(* IEC 61131-3 sources: daoli-st-library/DL_Process (part 18) *)

(* ---- FC_DL_TemperEmpiricalHardnessCalc.st ---- *)
(*
  Component : FC_DL_TemperEmpiricalHardnessCalc
  Category  : DL_Process
  Type      : FC
  Complexity: C2
  VERSION   : v1.0.0
  功能      : 回火温度-硬度经验曲线核算：按四点节点表分段线性插值得到基准 HRC，再按含碳量修正，超界双向钳位。
  开源溯源  : 道莅原创 clean-room 自研（无外部代码引用）｜License: MIT
  边界条件  : ① 节点表必须严格升序且首末温差 > 1e-9，否则返回哨兵 -1；
              ② 回火温度超出节点区间时取端点值并置 xClamped，禁外推；
              ③ 含碳量修正量双侧钳位 ±8 HRC，防小样本经验式发散。
*)
FUNCTION FC_DL_TemperEmpiricalHardnessCalc : REAL
VAR_INPUT
    fTemperC    : REAL;               (* 回火温度 [°C] Tempering temperature *)
    afTempKnot  : ARRAY[0..3] OF REAL;(* 节点温度表（升序） [°C] Knot temperatures ascending *)
    afHrcKnot   : ARRAY[0..3] OF REAL;(* 节点硬度表 [HRC] Knot hardness values *)
    fCarbonPct  : REAL;               (* 钢材含碳量 [%] Carbon content *)
END_VAR
VAR_OUTPUT
    fHrc      : REAL;   (* 插值得到的回火硬度 [HRC] Interpolated hardness *)
    fHrcCorr  : REAL;   (* 含碳量修正后的硬度 [HRC] Carbon-corrected hardness *)
    xClamped  : BOOL;   (* 超界钳位标志 [-] Out-of-range clamp flag *)
    xValid    : BOOL;   (* 计算有效性标志 [-] Calculation valid flag *)
END_VAR
VAR CONSTANT
    DL_EPS       : REAL := 1.0E-9;   (* 除零判定容差 [无量纲] Divide-by-zero tolerance *)
    DL_CORR_K    : REAL := 30.0;     (* 含碳量修正斜率 [HRC/%C] Carbon correction slope *)
    DL_CORR_BASE : REAL := 0.40;     (* 含碳量修正基准 [%C] Carbon correction base *)
    DL_CORR_LIM  : REAL := 8.0;      (* 含碳量修正钳位 [HRC] Carbon correction clamp *)
END_VAR
VAR
    nIdx  : INT;    (* 插值段循环下标 [-] Interpolation segment index *)
    nBad  : INT;    (* 节点表非有限计数，0 = 全部有限 [-] Non-finite knot counter *)
    fDen  : REAL;   (* 当前段温度跨度 [°C] Segment temperature span *)
    fCorr : REAL;   (* 含碳量修正量 [HRC] Carbon correction amount *)
END_VAR
(* 出口预置：四出口统一预置 *)
fHrc := 0.0; fHrcCorr := 0.0; xClamped := FALSE; xValid := FALSE; nBad := 0;
(* 非有限拦截：标量输入自反判 NaN，自身差值判 Inf *)
IF (fTemperC <> fTemperC) OR ((fTemperC - fTemperC) <> 0.0)
   OR (fCarbonPct <> fCarbonPct) OR ((fCarbonPct - fCarbonPct) <> 0.0) THEN
    FC_DL_TemperEmpiricalHardnessCalc := -1.0;  (* 哨兵 -1：输入非有限 / Sentinel -1 non-finite *)
    RETURN;
END_IF
(* 节点表非有限拦截：四个温度节点与四个硬度节点逐个判（越界读前先判界） *)
FOR nIdx := 0 TO 3 DO
    IF (nIdx >= 0) AND (nIdx <= 3) THEN
        IF (afTempKnot[nIdx] <> afTempKnot[nIdx])
           OR ((afTempKnot[nIdx] - afTempKnot[nIdx]) <> 0.0)
           OR (afHrcKnot[nIdx] <> afHrcKnot[nIdx])
           OR ((afHrcKnot[nIdx] - afHrcKnot[nIdx]) <> 0.0) THEN
            nBad := nBad + 1;
        END_IF
    END_IF
END_FOR
IF nBad > 0 THEN
    FC_DL_TemperEmpiricalHardnessCalc := -1.0;  (* 哨兵 -1：节点表非有限 / Sentinel -1 bad knots *)
    RETURN;
END_IF
(* 节点表域闸：首末温差必须为正，保证区间可插值与升序约定 *)
IF (afTempKnot[3] - afTempKnot[0]) <= DL_EPS THEN
    FC_DL_TemperEmpiricalHardnessCalc := -1.0;  (* 哨兵 -1：节点表非法 / Sentinel -1 bad knot table *)
    RETURN;
END_IF
(* 超界钳位：低于首节点取首值，高于末节点取末值，禁外推 *)
IF fTemperC <= afTempKnot[0] THEN
    fHrc := afHrcKnot[0];                       (* 端点取值 [HRC] / Lower endpoint *)
    xClamped := TRUE;                           (* 低位钳位标志 [-] / Low clamp *)
ELSIF fTemperC >= afTempKnot[3] THEN
    fHrc := afHrcKnot[3];                       (* 端点取值 [HRC] / Upper endpoint *)
    xClamped := TRUE;                           (* 高位钳位标志 [-] / High clamp *)
ELSE
    (* 分段线性插值：升序镜像遍历（禁倒序循环关键字），下标上限 2 保证 i+1 <= 3 不越界 *)
    FOR nIdx := 0 TO 2 DO
        IF (fTemperC >= afTempKnot[nIdx]) AND (fTemperC <= afTempKnot[nIdx + 1]) THEN
            fDen := afTempKnot[nIdx + 1] - afTempKnot[nIdx];   (* 段跨度 [°C] / Segment span *)
            IF ABS(fDen) > DL_EPS THEN
                fHrc := afHrcKnot[nIdx]
                        + (afHrcKnot[nIdx + 1] - afHrcKnot[nIdx])
                          * (fTemperC - afTempKnot[nIdx]) / fDen;
            END_IF
        END_IF
    END_FOR
END_IF
(* 含碳量修正：以 0.40 %C 为基准，每 0.1 %C 约 3 HRC，双侧钳位 *)
fCorr := (fCarbonPct - DL_CORR_BASE) * DL_CORR_K;
IF fCorr > DL_CORR_LIM THEN
    fCorr := DL_CORR_LIM;                       (* 上限钳位 [HRC] / Upper clamp *)
ELSIF fCorr < -DL_CORR_LIM THEN
    fCorr := -DL_CORR_LIM;                      (* 下限钳位 [HRC] / Lower clamp *)
END_IF
fHrcCorr := fHrc + fCorr;                       (* 修正后硬度 [HRC] / Corrected hardness *)
xValid := TRUE;                                 (* 链路有效 / Chain valid *)
FC_DL_TemperEmpiricalHardnessCalc := fHrcCorr;  (* 返回修正硬度 [HRC] / Return hardness *)
END_FUNCTION

(* ---- FC_DL_ThickenerSettlingAreaCalc.st ---- *)
(*
  Name: FC_DL_ThickenerSettlingAreaCalc
  Category: DL_Process
  Version: 1.0.0
  Round: R89 / 2026-11-25
  开源溯源：clean-room 自研（族 矿山破碎筛分，ST 开源生态实测 0 命中，无外部代码引入）
  功能：按固体体积衡算求浓密机底流体积流量与溢流量，再用沉降速度法算所需沉降面积与上升流速。
  边界条件：① 四入参全部过非有限闸，任一非有限返回哨兵 -1；
            ② 底流浓度必须显著高于给矿浓度（差值 ≥ 1 %），否则衡算无解，返回哨兵 -1；
            ③ 体积分数 φ 由质量分数与固/液密度反算，分母（固相项 + 液相项）在 0~1 质量分数域内恒正，
               仍以 DL_EPS 兜底防浮点下溢；面积取安全系数 1.15，上升流速 = Qo/A 故恒低于沉降速度。
  量纲自证：Q[m3/h] ÷ v[m/h] = m2；φ 无量纲。
*)
FUNCTION FC_DL_ThickenerSettlingAreaCalc : REAL
VAR_INPUT
    fFeedM3h : REAL;         (* 给矿浆体流量 [m3/h] Feed slurry flow [m3/h] *)
    fFeedSolidsPct : REAL;   (* 给矿固体质量浓度 [%] Feed solids mass concentration [%] *)
    fUnderSolidsPct : REAL;  (* 底流固体质量浓度 [%] Underflow solids mass concentration [%] *)
    fSettlingVel : REAL;     (* 自由沉降速度 [m/h] Free settling velocity [m/h] *)
END_VAR
VAR_OUTPUT
    fAreaM2 : REAL;          (* 所需沉降面积（含安全系数） [m2] Required settling area [m2] *)
    fRiseVel : REAL;         (* 溢流上升流速 [m/h] Overflow rise velocity [m/h] *)
    fOverflowM3h : REAL;     (* 溢流浆体流量 [m3/h] Overflow flow [m3/h] *)
    xSizingOk : BOOL;        (* 上升流速低于沉降速度则 TRUE [-] Rise velocity below settling velocity *)
    xValid : BOOL;           (* 计算有效性标志 [-] Calculation valid flag *)
END_VAR
VAR CONSTANT
    DL_EPS : REAL := 1.0E-9;      (* 除零判定容差 [-] Divide-by-zero tolerance *)
    DL_RHO_S : REAL := 2.7;       (* 固体密度（矿浆通用取值） [t/m3] Solids density [t/m3] *)
    DL_RHO_W : REAL := 1.0;       (* 液相密度（水） [t/m3] Liquid density [t/m3] *)
    DL_SF : REAL := 1.15;         (* 面积安全系数 [-] Area safety factor *)
    DL_PCT : REAL := 100.0;       (* 百分数基准 [%] Percent base *)
    DL_CONC_MIN_DIFF : REAL := 1.0; (* 底流与给矿浓度最小差值 [%] Minimum concentration difference *)
END_VAR
VAR
    fCf : REAL;     (* 给矿质量分数 [-] Feed mass fraction *)
    fCu : REAL;     (* 底流质量分数 [-] Underflow mass fraction *)
    fPhiF : REAL;   (* 给矿固体体积分数 [-] Feed solids volume fraction *)
    fPhiU : REAL;   (* 底流固体体积分数 [-] Underflow solids volume fraction *)
    fQs : REAL;     (* 固体体积流量 [m3/h] Solids volume flow [m3/h] *)
    fQu : REAL;     (* 底流浆体体积流量 [m3/h] Underflow slurry flow [m3/h] *)
    fQo : REAL;     (* 溢流浆体体积流量 [m3/h] Overflow flow [m3/h] *)
END_VAR
(* 出口预置：五出口统一预置（R256） *)
fAreaM2 := 0.0; fRiseVel := 0.0; fOverflowM3h := 0.0; xSizingOk := FALSE; xValid := FALSE;
(* 非有限闸：NaN 自反判 + Inf 差值自减判，四入参全枚举（R272） *)
IF (fFeedM3h <> fFeedM3h) OR ((fFeedM3h - fFeedM3h) <> 0.0)
   OR (fFeedSolidsPct <> fFeedSolidsPct) OR ((fFeedSolidsPct - fFeedSolidsPct) <> 0.0)
   OR (fUnderSolidsPct <> fUnderSolidsPct) OR ((fUnderSolidsPct - fUnderSolidsPct) <> 0.0)
   OR (fSettlingVel <> fSettlingVel) OR ((fSettlingVel - fSettlingVel) <> 0.0) THEN
    FC_DL_ThickenerSettlingAreaCalc := -1.0;    (* 哨兵 -1：入参非有限 / Sentinel -1, non-finite input *)
    RETURN;
END_IF
(* 组态域闸：流量与沉降速度为除子，浓度须物理可行且底流显著高于给矿 *)
IF (fFeedM3h <= DL_EPS) OR (fSettlingVel <= DL_EPS)
   OR (fFeedSolidsPct <= 0.0) OR (fFeedSolidsPct >= DL_PCT)
   OR (fUnderSolidsPct <= 0.0) OR (fUnderSolidsPct > DL_PCT)
   OR ((fUnderSolidsPct - fFeedSolidsPct) < DL_CONC_MIN_DIFF) THEN
    FC_DL_ThickenerSettlingAreaCalc := -1.0;    (* 哨兵 -1：组态非法 / Sentinel -1, bad configuration *)
    RETURN;
END_IF
fCf := fFeedSolidsPct / DL_PCT;                 (* 质量分数 [-] Mass fraction *)
fCu := fUnderSolidsPct / DL_PCT;
(* 体积分数：φ = (C/ρs) / (C/ρs + (1−C)/ρw)，固液体积可加性假设 *)
IF ((fCf / DL_RHO_S) + ((1.0 - fCf) / DL_RHO_W)) <= DL_EPS THEN
    FC_DL_ThickenerSettlingAreaCalc := -1.0;    (* 哨兵 -1：体积分数塌零 / Sentinel -1, vanishing phi *)
    RETURN;
END_IF
fPhiF := (fCf / DL_RHO_S) / ((fCf / DL_RHO_S) + ((1.0 - fCf) / DL_RHO_W));
fPhiU := (fCu / DL_RHO_S) / ((fCu / DL_RHO_S) + ((1.0 - fCu) / DL_RHO_W));
(* 固体体积衡算：Qs = Qf·φf；底流体积 Qu = Qs/φu，φu 已过域闸恒正 *)
IF fPhiU <= DL_EPS THEN
    FC_DL_ThickenerSettlingAreaCalc := -1.0;    (* 哨兵 -1：底流体积分数塌零 / Sentinel -1, phi underflow zero *)
    RETURN;
END_IF
fQs := fFeedM3h * fPhiF;                        (* 固体体积流量 [m3/h] Solids volume flow *)
fQu := fQs / fPhiU;                             (* 底流浆体流量 [m3/h] Underflow slurry flow *)
fQo := fFeedM3h - fQu;                          (* 溢流 = 给矿 − 底流 [m3/h] Overflow flow *)
IF fQo <= DL_EPS THEN
    FC_DL_ThickenerSettlingAreaCalc := -1.0;    (* 哨兵 -1：衡算无溢流，组态矛盾 / Sentinel -1, no overflow *)
    RETURN;
END_IF
(* 沉降面积：A = Qo/v × SF，Qo[m3/h] ÷ v[m/h] = m2 *)
fAreaM2 := (fQo / fSettlingVel) * DL_SF;
(* 上升流速：vR = Qo/A，A 已过正性检查（上式保证 ≥ SF 倍正量） *)
IF fAreaM2 <= DL_EPS THEN
    FC_DL_ThickenerSettlingAreaCalc := -1.0;    (* 哨兵 -1：面积塌零 / Sentinel -1, vanishing area *)
    RETURN;
END_IF
fRiseVel := fQo / fAreaM2;
fOverflowM3h := fQo;
(* 校核：上升流速低于自由沉降速度（含安全系数后恒成立，此处照实判定） *)
xSizingOk := fRiseVel < fSettlingVel;
xValid := TRUE;                                 (* 链路有效 / Chain valid *)
FC_DL_ThickenerSettlingAreaCalc := fAreaM2;
END_FUNCTION

(* ---- FC_DL_TinBathAtmosphereCalc.st ---- *)
(*
  Name: FC_DL_TinBathAtmosphereCalc
  Category: DL_Process
  Version: 1.0.0
  Round: R90 / 2026-11-25
  开源溯源：clean-room 自研（族 浮法玻璃锡槽退火，ST 开源生态实测 0 命中，无外部代码引入）
  功能：1) 锡槽保护气 H2 配比按「氢耗氧化学计量」估算。漏入锡槽的空气带入氧气，
           氧气与氢按 2H2 + O2 → 2H2O 反应，故 1 体积氧气需要 2 体积氢气中和。
           逐步为：
             氧带入量 = 漏入空气量 × 空气中氧体积分数(0.21)
             需中和氧量 = 氧带入量 − 允许残氧量（目标 ppm 折算为体积流量）
             氢需求 = 2 × 需中和氧量 × 过量系数
             氢配比 = 氢需求 / 保护气总流量 × 100
           允许残氧量按「目标 ppm × 总流量 × 1e-6」折算，使得目标越严格所需氢越多，方向正确。
        2) 过量系数 DL_HSF(1.5) 用于覆盖反应不完全与局部湍流死区，是安全冗余而非效率系数。
  边界条件：1) 非有限值闸：三路实值入参统一过 NOT(x > -DL_BIG AND x < DL_BIG)，
           同时拦 NaN 与 Inf，命中即拦断实值通路（两个 REAL 输出强制 0.0）并置无效（R19）。
        2) 分母零闸：ABS(fTotalFlowM3h) > DL_EPS 才允许算配比（总流量为 0 时配比无定义）。
        3) 负值闸：漏入量、目标氧含量、总流量任一为负判无效（不取绝对值掩盖反向）。
        4) 配比饱和钳制：H2 配比钳 0 ~ DL_H2_MAX(10 %)。上限的依据是保护气进入爆炸下限区间
           （H2 在空气中的爆炸下限约 4 %，但锡槽内为氮基气氛且需维持正压，工艺上按 10 % 上限组态），
           超过上限必须由安全联锁处理，本件只做钳制与无效标记，不做安全切断。
        5) 需求为负（残氧目标高于带入氧）时氢需求钳 0，属合法工况（无需加氢），不判无效。
        6) 饱和钳制：氢流量钳 0 ~ DL_H2_FLOW_MAX(10000 m3/h)，防溢出。
  量纲自证：氧带入量 = (m3/h) × [-] = m3/h；残氧量 = ppm × (m3/h) × 1E-6 = m3/h；
           需中和氧量 = (m3/h) − (m3/h) = m3/h，减法同量纲；
           氢需求 = [-] × (m3/h) × [-] = m3/h（化学计量比与过量系数均为无因次）；
           配比 = (m3/h) / (m3/h) × 100 = 无因次 [%]，分母与分子同量纲。
*)

FUNCTION FC_DL_TinBathAtmosphereCalc : BOOL
VAR_INPUT
    fO2TargetPpm   : REAL;   // 目标残氧含量 [ppm] / Target residual oxygen [ppm]
    fLeakM3h       : REAL;   // 漏入锡槽的空气量 [m3/h] / Air leakage into tin bath [m3/h]
    fTotalFlowM3h  : REAL;   // 保护气总流量 [m3/h] / Total protective gas flow [m3/h]
END_VAR
VAR_OUTPUT
    fH2Pct         : REAL;   // 氢气体积配比 [%] / Hydrogen volume ratio [%]
    fFlowM3h       : REAL;   // 氢气需求体积流量 [m3/h] / Hydrogen required volumetric flow [m3/h]
    xValid         : BOOL;   // 计算有效标志 [bool] / Calculation valid flag [bool]
END_VAR
VAR
    _fO2IngressM3h : REAL;   // 漏入氧气量 [m3/h] / Oxygen ingress [m3/h]
    _fO2AllowM3h   : REAL;   // 允许残氧量 [m3/h] / Allowable residual oxygen [m3/h]
    _fO2NeedM3h    : REAL;   // 需中和氧量 [m3/h] / Oxygen to be neutralized [m3/h]
    _fH2NeedM3h    : REAL;   // 氢需求（含过量系数）[m3/h] / Hydrogen demand with safety factor [m3/h]
    _fPctRaw       : REAL;   // 未饱和的配比 [%] / Raw ratio [%]
END_VAR
VAR CONSTANT
    DL_EPS         : REAL := 1.0E-9;    // 分母零闸阈值 [-] / Division-zero gate threshold [-]
    DL_BIG         : REAL := 1.0E12;    // 非有限值闸量级上限 [-] / Finiteness gate magnitude [-]
    DL_PCT         : REAL := 100.0;     // 百分比换算因子 [%] / Percent conversion factor [%]
    DL_O2_AIR_FRAC : REAL := 0.21;      // 空气中氧体积分数 [-] / Oxygen volume fraction in air [-]
    DL_H2_STOICH   : REAL := 2.0;       // 2H2 + O2 化学计量比 [-] / Hydrogen to oxygen stoichiometry [-]
    DL_PPM_FRAC    : REAL := 1.0E-6;    // ppm → 体积分数换算因子 [-] / ppm to volume fraction factor [-]
    DL_HSF         : REAL := 1.5;       // 氢过量系数（安全冗余）[-] / Hydrogen excess factor [-]
    DL_H2_MAX      : REAL := 10.0;      // 氢配比饱和上限 [%] / Hydrogen ratio saturation ceiling [%]
    DL_H2_FLOW_MAX : REAL := 10000.0;   // 氢流量饱和上限 [m3/h] / Hydrogen flow saturation ceiling [m3/h]
END_VAR

(* —— 段 1：非有限值闸（R19：三路入参全覆盖，拦 NaN 与 Inf） —— *)
IF NOT (fO2TargetPpm > -DL_BIG AND fO2TargetPpm < DL_BIG)
   OR NOT (fLeakM3h > -DL_BIG AND fLeakM3h < DL_BIG)
   OR NOT (fTotalFlowM3h > -DL_BIG AND fTotalFlowM3h < DL_BIG) THEN
    fH2Pct := 0.0;                          // 输出强制 0.0 / Output forced to zero
    fFlowM3h := 0.0;                        // 氢流量强制 0.0 / Hydrogen flow forced to zero
    xValid := FALSE;                        // 有效位清零 / Validity cleared
    FC_DL_TinBathAtmosphereCalc := FALSE;   // 返回码同源 / Return mirrors validity
    RETURN;                                 // 立即退出 / Immediate exit
END_IF

(* —— 段 2：分母零闸（R4：总流量是配比分母） —— *)
IF ABS(fTotalFlowM3h) <= DL_EPS THEN
    fH2Pct := 0.0;                          // 输出强制 0.0 / Output forced to zero
    fFlowM3h := 0.0;                        // 氢流量强制 0.0 / Hydrogen flow forced to zero
    xValid := FALSE;                        // 判无效 / Invalid
    FC_DL_TinBathAtmosphereCalc := FALSE;   // 返回码同步 / Return synchronised
    RETURN;                                 // 提前退出 / Early exit
END_IF

(* —— 段 3：负值闸（漏入量、目标氧含量、总流量均不可为负） —— *)
IF (fO2TargetPpm < 0.0) OR (fLeakM3h < 0.0) OR (fTotalFlowM3h < 0.0) THEN
    fH2Pct := 0.0;                          // 输出强制 0.0 / Output forced to zero
    fFlowM3h := 0.0;                        // 氢流量强制 0.0 / Hydrogen flow forced to zero
    xValid := FALSE;                        // 判无效 / Invalid
    FC_DL_TinBathAtmosphereCalc := FALSE;   // 返回码同步 / Return synchronised
    RETURN;                                 // 提前退出 / Early exit
END_IF

(* —— 段 4：氧衡算（R22 方向自核：漏入氧减去允许残氧，才是需要中和的量） —— *)
_fO2IngressM3h := fLeakM3h * DL_O2_AIR_FRAC;                      // 漏入氧气 [m3/h]
_fO2AllowM3h := fO2TargetPpm * DL_PPM_FRAC * fTotalFlowM3h;       // 允许残氧 [m3/h]
_fO2NeedM3h := MAX(0.0, _fO2IngressM3h - _fO2AllowM3h);           // 需中和氧量 [m3/h]（负值钳 0）

(* —— 段 5：氢需求与配比（化学计量比 2、过量系数 1.5 均为无因次） —— *)
_fH2NeedM3h := DL_H2_STOICH * _fO2NeedM3h * DL_HSF;               // 氢需求 [m3/h]
_fPctRaw := _fH2NeedM3h / fTotalFlowM3h * DL_PCT;                 // 氢配比 [%]

(* —— 段 6：输出单点写盘（饱和钳制） —— *)
fFlowM3h := LIMIT(0.0, _fH2NeedM3h, DL_H2_FLOW_MAX);              // 氢流量 [m3/h]
fH2Pct := LIMIT(0.0, _fPctRaw, DL_H2_MAX);                        // 氢配比 [%]

(* —— 段 7：有效位单点聚合（分母为正 + 入参非负） —— *)
xValid := (fTotalFlowM3h > DL_EPS)                                // 总流量为正
          AND (fO2TargetPpm >= 0.0)                               // 目标残氧非负
          AND (fLeakM3h >= 0.0);                                  // 漏入量非负
FC_DL_TinBathAtmosphereCalc := xValid;                            // 返回码：TRUE = 计算可信

END_FUNCTION

(* ---- FC_DL_TireCureBladderSteamCalc.st ---- *)
(*
  Name: FC_DL_TireCureBladderSteamCalc
  Category: DL_Process
  Version: 1.0.0
  Round: R91 / 2026-11-25
  开源溯源：clean-room 自研（族 轮胎硫化，ST 开源生态实测 0 命中，无外部代码引入）
  功能：1) 单周期胶囊蒸汽耗量按「充装量 + 升温量 + 排凝损失」三段求和：
           充装量 = 胶囊容积 * 蒸汽密度；
           升温量 = 胶囊内容物质量 * 比热 * 温升 / 潜热（把显热需求折成蒸汽质量）；
           排凝损失 = (充装量 + 升温量) * fDrainPct / 100。
           即 m = (V*rho + m*cp*dT/hfg) * (1 + drainPct/100)，单位 kg/周期。
        2) 输出分解量 fFillKg 与 fHeatUpKg，便于按段归因能耗（充装段与升温段的节能措施完全不同）。
        3) 容积零闸与潜热零闸：胶囊容积为充装量的乘子、潜热为升温量的分母，
           任一为零会把「未组态」伪装成「零耗量」，必须判无效而非输出 0。
  边界条件：1) 非有限值闸：七路实值入参先过 NOT(x > -DL_BIG AND x < DL_BIG)，同时拦 NaN 与 Inf，
           命中即闸断实值通路（三段耗量与总耗量强制 0.0），不得只置标志（R19）。
        2) 分母零闸：升华/汽化潜热 fLatentKjKg 必须 > DL_EPS；胶囊内容物比热 fWaterCpKjKgK 必须 > DL_EPS。
        3) 容积零闸：fBladderVolL 必须 > DL_EPS；蒸汽密度 fSteamDensityKgm3 必须 > DL_EPS。
        4) 排凝率域闸：fDrainPct 必须落在 [0.0, DL_DRAIN_HI] 内（排凝率超 100 % 不具物理意义），
           越域判无效不钳制。
        5) 判据取原始值（R24）：总量越域判定使用钳制前的 _fTotalRawKg，钳制只作用于输出。
        6) 纯函数无状态：单周期耗量的累计与班产统计由上层计量模块承担。
  量纲自证：V [L] * rho [kg/m3] / 1000 [L/m3] = kg；
           m [kg] * cp [kJ/(kg*K)] * dT [K] = kJ；kJ / hfg [kJ/kg] = kg；
           三段同为 kg，求和合法；排凝率为无因次百分数，乘 kg 仍为 kg。
  修订历史 Revision :
    2026-11-25  v1.0.0  R91 首版
*)

FUNCTION FC_DL_TireCureBladderSteamCalc : BOOL
VAR_INPUT
    fBladderVolL     : REAL;   // 胶囊有效容积 [L] / Effective bladder volume [L]
    fSteamDensityKgm3 : REAL;  // 工作压力下蒸汽密度 [kg/m3] / Steam density at working pressure [kg/m3]
    fContentMassKg   : REAL;   // 胶囊内容物（水/氮）质量 [kg] / Bladder content mass [kg]
    fWaterCpKjKgK    : REAL;   // 内容物比热 [kJ/(kg*K)] / Content specific heat [kJ/(kg*K)]
    fTempRiseK       : REAL;   // 升温幅度 [K] / Temperature rise [K]
    fLatentKjKg      : REAL;   // 工作压力下汽化潜热 [kJ/kg] / Latent heat of vaporisation [kJ/kg]
    fDrainPct        : REAL;   // 排凝损失占充装与升温之和的百分比 [%] / Blowdown loss percentage [%]
END_VAR
VAR_OUTPUT
    fFillKg          : REAL;   // 充装段蒸汽量 [kg] / Steam for initial filling [kg]
    fHeatUpKg        : REAL;   // 升温段蒸汽量 [kg] / Steam for heat-up [kg]
    fSteamKg         : REAL;   // 单周期蒸汽总耗量 [kg/cycle] / Total steam consumption per cycle [kg/cycle]
    xValid           : BOOL;   // 计算有效标志 [bool] / Calculation valid flag [bool]
END_VAR
VAR
    _fFillRawKg      : REAL;   // 钳制前的充装量 [kg] / Raw fill mass [kg]
    _fHeatRawKg      : REAL;   // 钳制前的升温量 [kg] / Raw heat-up mass [kg]
    _fTotalRawKg     : REAL;   // 钳制前的总量 [kg] / Raw total mass [kg]
    _fDrainFactor    : REAL;   // 排凝放大因子（1 + 排凝率/100）[-] / Blowdown multiplier [-]
END_VAR
VAR CONSTANT
    DL_EPS           : REAL := 1.0E-9;    // 数值零闸阈值 [-] / Numeric zero gate threshold [-]
    DL_BIG           : REAL := 1.0E12;    // 非有限值闸量级上限 [-] / Finiteness gate magnitude [-]
    DL_L_PER_M3      : REAL := 1000.0;    // 立方米到升的折算 [L/m3] / Litres per cubic metre [L/m3]
    DL_PCT           : REAL := 100.0;     // 百分比换算因子 [%] / Percent conversion factor [%]
    DL_DRAIN_HI      : REAL := 100.0;     // 排凝率物理上限 [%] / Blowdown percentage upper bound [%]
    DL_STEAM_HI_KG   : REAL := 5000.0;    // 单周期耗量物理上限 [kg] / Steam mass physical upper bound [kg]
END_VAR

(* —— 段 1：非有限值闸（R19：闸断实值通路） —— *)
IF NOT (fBladderVolL > -DL_BIG AND fBladderVolL < DL_BIG)
   OR NOT (fSteamDensityKgm3 > -DL_BIG AND fSteamDensityKgm3 < DL_BIG)
   OR NOT (fContentMassKg > -DL_BIG AND fContentMassKg < DL_BIG)
   OR NOT (fWaterCpKjKgK > -DL_BIG AND fWaterCpKjKgK < DL_BIG)
   OR NOT (fTempRiseK > -DL_BIG AND fTempRiseK < DL_BIG)
   OR NOT (fLatentKjKg > -DL_BIG AND fLatentKjKg < DL_BIG)
   OR NOT (fDrainPct > -DL_BIG AND fDrainPct < DL_BIG) THEN
    fFillKg := 0.0;                         // 充装量强制 0.0 / Fill mass forced to zero
    fHeatUpKg := 0.0;                       // 升温量强制 0.0 / Heat-up mass forced to zero
    fSteamKg := 0.0;                        // 总量强制 0.0，切断污染源 / Total forced to zero
    xValid := FALSE;                        // 有效位清零 / Validity cleared
    FC_DL_TireCureBladderSteamCalc := FALSE;   // 返回码与有效位同源 / Return mirrors validity
    RETURN;                                 // 立即退出 / Immediate exit
END_IF

(* —— 段 2：分母零闸与域闸（容积/密度为乘子，潜热/比热为分母） —— *)
IF (fBladderVolL <= DL_EPS)                                       // 容积不可为零
   OR (fSteamDensityKgm3 <= DL_EPS)                               // 蒸汽密度不可为零
   OR (fContentMassKg < 0.0)                                      // 内容物质量不得为负
   OR (fWaterCpKjKgK <= DL_EPS)                                   // 比热不可为零
   OR (fTempRiseK < 0.0)                                          // 升温幅度不得为负（方向固定）
   OR (fLatentKjKg <= DL_EPS)                                     // 潜热不可为零
   OR (fDrainPct < 0.0)                                           // 排凝率不得为负
   OR (fDrainPct > DL_DRAIN_HI) THEN                              // 排凝率不得超 100 %
    fFillKg := 0.0;                         // 参数不可用即无耗量 / No parameter, no consumption
    fHeatUpKg := 0.0;                       // 升温量不可算 / Heat-up mass not computable
    fSteamKg := 0.0;                        // 总量不可算 / Total not computable
    xValid := FALSE;                        // 判无效 / Invalid
    FC_DL_TireCureBladderSteamCalc := FALSE;   // 返回码同步 / Return synchronised
    RETURN;                                 // 提前退出 / Early exit
END_IF

(* —— 段 3：主算式（不钳制，先出原始值供段 4 判据使用，R24） —— *)
_fFillRawKg := fBladderVolL / DL_L_PER_M3 * fSteamDensityKgm3;                     // 充装段 [kg]
_fHeatRawKg := fContentMassKg * fWaterCpKjKgK * fTempRiseK / fLatentKjKg;          // 升温段折蒸汽 [kg]
_fDrainFactor := 1.0 + fDrainPct / DL_PCT;                                        // 排凝放大因子 [-]
_fTotalRawKg := (_fFillRawKg + _fHeatRawKg) * _fDrainFactor;                       // 单周期总量 [kg]

(* —— 段 4：判据（取原始值；单点 BOOL 聚合避免多处赋 FALSE 覆盖） —— *)
xValid := (_fFillRawKg >= 0.0)                                                    // 充装量不得为负
          AND (_fHeatRawKg >= 0.0)                                                // 升温量不得为负
          AND (_fTotalRawKg >= 0.0)                                               // 总量不得为负
          AND (_fTotalRawKg <= DL_STEAM_HI_KG);                                   // 不得超物理上限（量级异常）

(* —— 段 5：输出单点写盘（钳制到物理域内，判定结果已在段 4 定案） —— *)
fFillKg := LIMIT(0.0, _fFillRawKg, DL_STEAM_HI_KG);                               // 充装段钳物理域 [kg]
fHeatUpKg := LIMIT(0.0, _fHeatRawKg, DL_STEAM_HI_KG);                             // 升温段钳物理域 [kg]
fSteamKg := LIMIT(0.0, _fTotalRawKg, DL_STEAM_HI_KG);                             // 总量钳物理域 [kg/cycle]
FC_DL_TireCureBladderSteamCalc := xValid;                                         // 返回码：TRUE = 计算可信

END_FUNCTION

(* ---- FC_DL_TireCureDegreeCalc.st ---- *)
(*
  Name: FC_DL_TireCureDegreeCalc
  Category: DL_Process
  Version: 1.0.0
  Round: R91 / 2026-11-25
  开源溯源：clean-room 自研（族 轮胎硫化，ST 开源生态实测 0 命中，无外部代码引入）
  功能：1) 硫化程度按「实际等效硫化时间 / 目标等效硫化时间」计算并折百分比：
           degree = t_equiv / t_target * 100，其中 t_equiv 由 FC_DL_TireCureEquivalentTimeCalc
           给出的 140 degC 基准当量时间（本件不重复其换算，只做比值判据，故本件仍自包含无依赖）。
        2) 欠硫 / 过硫判定：degree < fUnderPct 判欠硫（物理性能不达标，须延长硫化）；
           degree > fOverPct 判过硫（返原、断裂伸长下降，须缩短硫化或降低模温）。
           两个阈值各占一个独立布尔出口，供上层分别处置（欠硫可补救，过硫不可逆）。
        3) 输出硫化程度百分比同时钳到 [0.0, DL_DEG_HI]（DL_DEG_HI = 200 %），
           保留超硫观测余量的同时避免极端值污染趋势曲线。
  边界条件：1) 非有限值闸：四路实值入参先过 NOT(x > -DL_BIG AND x < DL_BIG)，同时拦 NaN 与 Inf，
           命中即闸断实值通路（程度强制 0.0 且置欠硫位，保守侧），不得只置标志（R19）。
        2) 分母零闸：目标等效时间 fTargetEquivMin 必须 > DL_EPS（比值式分母），
           否则判无效并清零 —— 输出「未组态即 0 %」会被误读为「完全没有硫化」。
        3) 阈值域闸：须满足 0.0 < fUnderPct < fOverPct <= DL_DEG_HI，否则两级判据重叠或倒置，
           越域判无效并把欠硫位置真（保守侧）。
        4) 时间非负闸：实际等效时间不得为负（负值属积分方向错误），判无效。
        5) 判据取原始值（R24）：欠硫/过硫判定使用钳制前的 _fDegreeRawPct，不得先钳再判。
        6) 纯函数无状态：等效时间本身的积分与累计由上层硫化序 FB 承担。
  量纲自证：degree = (min)/(min)*100 = 无因次百分数 [%]；
           fUnderPct / fOverPct 同为百分数，可与 degree 直接比较，量纲合法。
  修订历史 Revision :
    2026-11-25  v1.0.0  R91 首版
*)

FUNCTION FC_DL_TireCureDegreeCalc : BOOL
VAR_INPUT
    fEquivTimeMin    : REAL;   // 实际等效硫化时间（140 degC 基准）[min] / Actual equivalent cure time [min]
    fTargetEquivMin  : REAL;   // 目标等效硫化时间 [min] / Target equivalent cure time [min]
    fUnderPct        : REAL;   // 欠硫判定阈值 [%] / Under-cure threshold [%]
    fOverPct         : REAL;   // 过硫判定阈值 [%] / Over-cure threshold [%]
END_VAR
VAR_OUTPUT
    fDegreePct       : REAL;   // 硫化程度 [%] / Degree of cure [%]
    xUnderCure       : BOOL;   // 欠硫标志 [bool] / Under-cure flag [bool]
    xOverCure        : BOOL;   // 过硫标志 [bool] / Over-cure flag [bool]
    xValid           : BOOL;   // 计算有效标志 [bool] / Calculation valid flag [bool]
END_VAR
VAR
    _fDegreeRawPct   : REAL;   // 钳制前的原始硫化程度 [%] / Raw degree of cure before limiting [%]
END_VAR
VAR CONSTANT
    DL_EPS           : REAL := 1.0E-9;    // 数值零闸阈值 [-] / Numeric zero gate threshold [-]
    DL_BIG           : REAL := 1.0E12;    // 非有限值闸量级上限 [-] / Finiteness gate magnitude [-]
    DL_PCT           : REAL := 100.0;     // 百分比换算因子 [%] / Percent conversion factor [%]
    DL_DEG_HI        : REAL := 200.0;     // 硫化程度显示上限（留过硫观测余量）[%] / Degree display ceiling [%]
    DL_ZERO_PCT      : REAL := 0.0;       // 百分数零基准 [%] / Zero percent reference [%]
END_VAR

(* —— 段 1：非有限值闸（R19：闸断实值通路；失效侧置欠硫位，保守侧） —— *)
IF NOT (fEquivTimeMin > -DL_BIG AND fEquivTimeMin < DL_BIG)
   OR NOT (fTargetEquivMin > -DL_BIG AND fTargetEquivMin < DL_BIG)
   OR NOT (fUnderPct > -DL_BIG AND fUnderPct < DL_BIG)
   OR NOT (fOverPct > -DL_BIG AND fOverPct < DL_BIG) THEN
    fDegreePct := 0.0;                      // 输出强制 0.0，切断污染源 / Force zero, cut polluted path
    xUnderCure := TRUE;                     // 失效侧按欠硫处理（保守侧：宁可延长不可放行）
    xOverCure := FALSE;                     // 失效侧过硫位保持假 / Over-cure stays false
    xValid := FALSE;                        // 有效位清零 / Validity cleared
    FC_DL_TireCureDegreeCalc := FALSE;      // 返回码与有效位同源 / Return mirrors validity
    RETURN;                                 // 立即退出 / Immediate exit
END_IF

(* —— 段 2：分母零闸与阈值域闸（目标时间为比值分母） —— *)
IF (fTargetEquivMin <= DL_EPS)                                    // 目标时间不可为零
   OR (fEquivTimeMin < 0.0)                                       // 实际时间不得为负
   OR (fUnderPct <= DL_ZERO_PCT)                                  // 欠硫阈值必须为正
   OR (fOverPct <= fUnderPct)                                     // 过硫阈值必须大于欠硫阈值
   OR (fOverPct > DL_DEG_HI) THEN                                 // 过硫阈值不得超显示上限
    fDegreePct := 0.0;                      // 参数不可用即无程度 / No parameter, no degree
    xUnderCure := TRUE;                     // 按欠硫处理（保守侧）/ Treat as under-cured
    xOverCure := FALSE;                     // 过硫位保持假 / Over-cure stays false
    xValid := FALSE;                        // 判无效 / Invalid
    FC_DL_TireCureDegreeCalc := FALSE;      // 返回码同步 / Return synchronised
    RETURN;                                 // 提前退出 / Early exit
END_IF

(* —— 段 3：主算式（不钳制，先出原始值供段 4 判据使用，R24） —— *)
_fDegreeRawPct := fEquivTimeMin / fTargetEquivMin * DL_PCT;                       // 硫化程度 [%]

(* —— 段 4：判据（取原始值；单点 BOOL 聚合避免多处赋 FALSE 覆盖） —— *)
xUnderCure := (_fDegreeRawPct < fUnderPct);                                       // 欠硫
xOverCure := (_fDegreeRawPct > fOverPct);                                         // 过硫
xValid := (_fDegreeRawPct >= DL_ZERO_PCT)                                         // 程度不得为负（方向固定）
          AND (_fDegreeRawPct <= DL_DEG_HI);                                      // 不得超显示上限（量级异常）

(* —— 段 5：输出单点写盘（钳制到显示域内，判定结果已在段 4 定案） —— *)
fDegreePct := LIMIT(DL_ZERO_PCT, _fDegreeRawPct, DL_DEG_HI);                      // 程度钳 0..200 [%]
FC_DL_TireCureDegreeCalc := xValid;                                               // 返回码：TRUE = 计算可信

END_FUNCTION

(* ---- FC_DL_TireCureEquivalentTimeCalc.st ---- *)
(*
  Name: FC_DL_TireCureEquivalentTimeCalc
  Category: DL_Process
  Version: 1.0.0
  Round: R91 / 2026-11-25
  开源溯源：clean-room 自研（族 轮胎硫化，ST 开源生态实测 0 命中，无外部代码引入）
  功能：1) 等效硫化时间按 Arrhenius 温度-时间等效原理折算到 140 degC 基准：
           速率比 R = EXP( (Ea/Rg) * (1/T_ref − 1/T_cur) )，
           t_eq = t_cur * R，其中 T 一律换算为绝对温度 [K]，Ea 为表观活化能 [J/mol]，
           Rg 为通用气体常数 8.314 [J/(mol*K)]；温度高于基准时 R > 1（硫化更快）。
        2) 输出两个量：等效时间 fEquivTimeMin [min] 与速率比 fRateRatio [-]，
           后者便于观察当前温度折算强度（R = 2 表示 1 min 相当于基准温度的 2 min）。
        3) 温度域校验：当前温度与基准温度都必须高于绝对零度（换算后 T > 0 K），
           否则 1/T 无意义；越域判无效并清零全部输出，绝不让除零结果流到下游。
  边界条件：1) 非有限值闸：四路实值入参先过 NOT(x > -DL_BIG AND x < DL_BIG)，同时拦 NaN 与 Inf，
           命中即闸断实值通路（等效时间与速率比强制 0.0），不得只置标志（R19）。
        2) 温度零闸：开尔文换算后 T_cur / T_ref 必须 > DL_T_K_MIN（取 1.0 K 作下限，
           远高于绝对零度，同时拦住「传摄氏值当开尔文」的组态错），否则判无效。
        3) 活化能域闸：fActEnergyKjMol 必须落在 (DL_EA_LO, DL_EA_HI) 内 ——
           橡胶硫化表观活化能工程带约 80 ~ 200 kJ/mol，越域说明单位用错（J 与 kJ 混用）。
        4) 指数溢出闸：指数 = (Ea/Rg)*(1/Tref − 1/Tcur)，在合法温度域内其绝对值有界；
           仍显式钳制到 [-DL_EXPO_HI, +DL_EXPO_HI]，防 EXP 溢出为 Inf 后穿透（R19 第二道）。
        5) 判据取原始值（R24）：等效时间越域判定使用钳制前的 _fEquivRawMin，钳制只作用于输出。
        6) 纯函数无状态：温度积分的累计由硫化程度件（FC_DL_TireCureDegreeCalc）承担。
  量纲自证：(Ea/Rg) = (J/mol)/(J/(mol*K)) = K；乘 (1/K − 1/K) = 1/K 得无因次，故 EXP 自变量无因次；
           t_eq = (min) * (无因次) = min，与 fRefTimeMin 同量纲。
  修订历史 Revision :
    2026-11-25  v1.0.0  R91 首版
*)

FUNCTION FC_DL_TireCureEquivalentTimeCalc : BOOL
VAR_INPUT
    fCureTempC       : REAL;   // 当前硫化温度 [degC] / Current curing temperature [degC]
    fCureTimeMin     : REAL;   // 当前温度下的实际硫化时间 [min] / Actual curing time at current temperature [min]
    fActEnergyKjMol  : REAL;   // 表观活化能 [kJ/mol] / Apparent activation energy [kJ/mol]
    fRefTempC        : REAL;   // 等效基准温度（通常 140 degC）[degC] / Reference temperature, usually 140 degC [degC]
    fRefTimeMin      : REAL;   // 基准温度下的标准硫化时间 [min] / Standard cure time at reference temperature [min]
END_VAR
VAR_OUTPUT
    fEquivTimeMin    : REAL;   // 折算后的等效硫化时间 [min] / Equivalent curing time at reference temperature [min]
    fRateRatio       : REAL;   // 速率比（当前温度相对基准）[-] / Rate ratio against the reference [-]
    xValid           : BOOL;   // 计算有效标志 [bool] / Calculation valid flag [bool]
END_VAR
VAR
    _fCurK           : REAL;   // 当前绝对温度 [K] / Current absolute temperature [K]
    _fRefK           : REAL;   // 基准绝对温度 [K] / Reference absolute temperature [K]
    _fEaJmol         : REAL;   // 表观活化能 [J/mol] / Apparent activation energy [J/mol]
    _fExpo           : REAL;   // Arrhenius 指数（无因次）[-] / Arrhenius exponent, dimensionless [-]
    _fRatioRaw       : REAL;   // 未钳制的速率比 [-]/ Unclamped rate ratio [-]
    _fEquivRawMin    : REAL;   // 钳制前的等效时间 [min] / Raw equivalent time before limiting [min]
END_VAR
VAR CONSTANT
    DL_EPS           : REAL := 1.0E-9;    // 数值零闸阈值 [-] / Numeric zero gate threshold [-]
    DL_BIG           : REAL := 1.0E12;    // 非有限值闸量级上限 [-] / Finiteness gate magnitude [-]
    DL_KELVIN_OFF    : REAL := 273.15;    // 摄氏到开尔文的偏移 [K] / Celsius to Kelvin offset [K]
    DL_T_K_MIN       : REAL := 1.0;       // 绝对温度下限（护栏）[K] / Absolute temperature floor [K]
    DL_EA_LO         : REAL := 50.0;      // 硫化表观活化能域下限 [kJ/mol] / Activation energy domain low [kJ/mol]
    DL_EA_HI         : REAL := 300.0;     // 硫化表观活化能域上限 [kJ/mol] / Activation energy domain high [kJ/mol]
    DL_J_PER_KJ      : REAL := 1000.0;    // 千焦到焦的折算 [J/kJ] / Joules per kilojoule [J/kJ]
    DL_RG            : REAL := 8.314;     // 通用气体常数 [J/(mol*K)] / Universal gas constant [J/(mol*K)]
    DL_EXPO_HI       : REAL := 50.0;      // 指数钳制上限（防 EXP 溢出）[-] / Exponent clamp bound against overflow [-]
    DL_TIME_HI_MIN   : REAL := 100000.0;  // 等效时间物理上限 [min] / Equivalent time physical upper bound [min]
END_VAR

(* —— 段 1：非有限值闸（R19：闸断实值通路） —— *)
IF NOT (fCureTempC > -DL_BIG AND fCureTempC < DL_BIG)
   OR NOT (fCureTimeMin > -DL_BIG AND fCureTimeMin < DL_BIG)
   OR NOT (fActEnergyKjMol > -DL_BIG AND fActEnergyKjMol < DL_BIG)
   OR NOT (fRefTempC > -DL_BIG AND fRefTempC < DL_BIG)
   OR NOT (fRefTimeMin > -DL_BIG AND fRefTimeMin < DL_BIG) THEN
    fEquivTimeMin := 0.0;                   // 输出强制 0.0，切断污染源 / Force zero, cut polluted path
    fRateRatio := 0.0;                      // 速率比强制 0.0 / Rate ratio forced to zero
    xValid := FALSE;                        // 有效位清零 / Validity cleared
    FC_DL_TireCureEquivalentTimeCalc := FALSE;   // 返回码与有效位同源 / Return mirrors validity
    RETURN;                                 // 立即退出 / Immediate exit
END_IF

(* —— 段 2：温度零闸（绝对温度必须为正，否则 1/T 无意义） —— *)
_fCurK := fCureTempC + DL_KELVIN_OFF;                                     // 当前绝对温度 [K]
_fRefK := fRefTempC + DL_KELVIN_OFF;                                      // 基准绝对温度 [K]
IF (_fCurK <= DL_T_K_MIN) OR (_fRefK <= DL_T_K_MIN) THEN
    fEquivTimeMin := 0.0;                   // 温度越域即不可算 / Temperature out of domain
    fRateRatio := 0.0;                      // 速率比不可算 / Rate ratio not computable
    xValid := FALSE;                        // 判无效 / Invalid
    FC_DL_TireCureEquivalentTimeCalc := FALSE;   // 返回码同步 / Return synchronised
    RETURN;                                 // 提前退出 / Early exit
END_IF

(* —— 段 3：活化能域闸（防 J 与 kJ 单位混用） —— *)
IF (fActEnergyKjMol <= DL_EA_LO) OR (fActEnergyKjMol >= DL_EA_HI) THEN
    fEquivTimeMin := 0.0;                   // 活化能越域即不可算 / Activation energy out of domain
    fRateRatio := 0.0;                      // 速率比不可算 / Rate ratio not computable
    xValid := FALSE;                        // 判无效 / Invalid
    FC_DL_TireCureEquivalentTimeCalc := FALSE;   // 返回码同步 / Return synchronised
    RETURN;                                 // 提前退出 / Early exit
END_IF

(* —— 段 4：主算式（指数先钳制再 EXP，防溢出为 Inf 穿透） —— *)
_fEaJmol := fActEnergyKjMol * DL_J_PER_KJ;                                        // 活化能 [J/mol]
_fExpo := _fEaJmol / DL_RG * (1.0 / _fRefK - 1.0 / _fCurK);                       // Arrhenius 指数 [-]
_fExpo := LIMIT(-DL_EXPO_HI, _fExpo, DL_EXPO_HI);                                 // 指数钳制（第二道溢出闸）
_fRatioRaw := EXP(_fExpo);                                                        // 速率比 [-]
_fEquivRawMin := fCureTimeMin * _fRatioRaw;                                       // 等效时间 [min]

(* —— 段 5：判据（取原始值；单点 BOOL 聚合避免多处赋 FALSE 覆盖） —— *)
xValid := (fCureTimeMin >= 0.0)                                                   // 时间不得为负
          AND (fRefTimeMin > 0.0)                                                 // 基准时间必须为正
          AND (_fRatioRaw > 0.0)                                                  // 速率比必须为正（EXP 恒正）
          AND (_fEquivRawMin >= 0.0)                                              // 等效时间不得为负
          AND (_fEquivRawMin <= DL_TIME_HI_MIN);                                  // 不得超物理上限（量级异常）

(* —— 段 6：输出单点写盘（钳制到物理域内，判定结果已在段 5 定案） —— *)
fEquivTimeMin := LIMIT(0.0, _fEquivRawMin, DL_TIME_HI_MIN);                       // 等效时间钳物理域 [min]
fRateRatio := _fRatioRaw;                                                         // 速率比出口（恒正，无需钳负侧）
FC_DL_TireCureEquivalentTimeCalc := xValid;                                       // 返回码：TRUE = 计算可信

END_FUNCTION

(* ---- FC_DL_TireCureMoldCycleTimeCalc.st ---- *)
(*
  Name: FC_DL_TireCureMoldCycleTimeCalc
  Category: DL_Process
  Version: 1.0.0
  Round: R91 / 2026-11-25
  开源溯源：clean-room 自研（族 轮胎硫化，ST 开源生态实测 0 命中，无外部代码引入）
  功能：1) 模压周期按「合模 + 升温 + 保温 + 排凝 + 开模」五段求和：
           fCycleMin = tClose + tHeat + tHold + tBlowDown + tOpen，各段以分钟给出，同量纲直加。
        2) 输出保温段占比 fHoldSharePct = tHold / 总周期 * 100，用于判断周期结构是否合理
           （硫化周期的绝大部分应为保温段；保温占比过低意味着辅助动作时间过长、机台利用率差）。
        3) 分段零值容错：允许任一段为 0（例如无排凝动作的机台把 tBlowDown 组态为 0），
           但总周期必须 > DL_EPS，否则「零周期」无法作为节拍基准，判无效。
  边界条件：1) 非有限值闸：五路实值入参先过 NOT(x > -DL_BIG AND x < DL_BIG)，同时拦 NaN 与 Inf，
           命中即闸断实值通路（总周期与占比强制 0.0），不得只置标志（R19）。
        2) 分段非负闸：任一段为负即判无效（负时长属组态错，求和时会被掩盖成「周期偏短」），
           绝不取绝对值或按 0 处理。
        3) 总周期零闸：总周期 <= DL_EPS 时占比式分母为零，判无效并清零，不输出无穷大占比。
        4) 分段上限闸：单段超过 DL_SEG_HI_MIN（12 小时）判无效 —— 超过整模寿命量级的组态
           几乎必然是单位用错（秒当作分）。
        5) 判据取原始值（R24）：总周期与占比越域判定均使用钳制前的原始值，不先钳后判。
        6) 物理域钳制：总周期钳 0.0 ~ DL_CYCLE_HI_MIN；占比钳 0.0 ~ DL_PCT_HI。
  量纲自证：五段均为 [min]，直加得 [min]；
           fHoldSharePct = (min)/(min)*100 = 无因次百分数 [%]，量纲合法。
  修订历史 Revision :
    2026-11-25  v1.0.0  R91 首版
*)

FUNCTION FC_DL_TireCureMoldCycleTimeCalc : BOOL
VAR_INPUT
    fCloseMin        : REAL;   // 合模段时长 [min] / Mold closing segment duration [min]
    fHeatMin         : REAL;   // 升温段时长 [min] / Heat-up segment duration [min]
    fHoldMin         : REAL;   // 保温（硫化）段时长 [min] / Curing hold segment duration [min]
    fBlowDownMin     : REAL;   // 排凝段时长 [min] / Blowdown segment duration [min]
    fOpenMin         : REAL;   // 开模段时长 [min] / Mold opening segment duration [min]
END_VAR
VAR_OUTPUT
    fCycleMin        : REAL;   // 模压周期总时长 [min] / Total mold cycle time [min]
    fHoldSharePct    : REAL;   // 保温段占周期百分比 [%] / Hold segment share of the cycle [%]
    xValid           : BOOL;   // 计算有效标志 [bool] / Calculation valid flag [bool]
END_VAR
VAR
    _fCycleRawMin    : REAL;   // 钳制前的原始总周期 [min] / Raw total cycle before limiting [min]
    _fShareRawPct    : REAL;   // 钳制前的原始占比 [%] / Raw share before limiting [%]
END_VAR
VAR CONSTANT
    DL_EPS           : REAL := 1.0E-9;    // 数值零闸阈值 [-] / Numeric zero gate threshold [-]
    DL_BIG           : REAL := 1.0E12;    // 非有限值闸量级上限 [-] / Finiteness gate magnitude [-]
    DL_PCT           : REAL := 100.0;     // 百分比换算因子 [%] / Percent conversion factor [%]
    DL_PCT_HI        : REAL := 100.0;     // 占比物理上限 [%] / Share upper bound [%]
    DL_SEG_HI_MIN    : REAL := 720.0;     // 单段时长上限（12 小时）[min] / Single segment upper bound, 12 h [min]
    DL_CYCLE_HI_MIN  : REAL := 720.0;     // 总周期物理上限 [min] / Total cycle physical upper bound [min]
END_VAR

(* —— 段 1：非有限值闸（R19：闸断实值通路） —— *)
IF NOT (fCloseMin > -DL_BIG AND fCloseMin < DL_BIG)
   OR NOT (fHeatMin > -DL_BIG AND fHeatMin < DL_BIG)
   OR NOT (fHoldMin > -DL_BIG AND fHoldMin < DL_BIG)
   OR NOT (fBlowDownMin > -DL_BIG AND fBlowDownMin < DL_BIG)
   OR NOT (fOpenMin > -DL_BIG AND fOpenMin < DL_BIG) THEN
    fCycleMin := 0.0;                       // 输出强制 0.0，切断污染源 / Force zero, cut polluted path
    fHoldSharePct := 0.0;                   // 占比强制 0.0 / Share forced to zero
    xValid := FALSE;                        // 有效位清零 / Validity cleared
    FC_DL_TireCureMoldCycleTimeCalc := FALSE;   // 返回码与有效位同源 / Return mirrors validity
    RETURN;                                 // 立即退出 / Immediate exit
END_IF

(* —— 段 2：分段非负闸与上限闸（负时长会把周期掩盖成偏短，必须判无效） —— *)
IF (fCloseMin < 0.0) OR (fHeatMin < 0.0) OR (fHoldMin < 0.0)
   OR (fBlowDownMin < 0.0) OR (fOpenMin < 0.0) THEN
    fCycleMin := 0.0;                       // 负时长即不可算 / Negative duration is not computable
    fHoldSharePct := 0.0;                   // 占比不可算 / Share not computable
    xValid := FALSE;                        // 判无效 / Invalid
    FC_DL_TireCureMoldCycleTimeCalc := FALSE;   // 返回码同步 / Return synchronised
    RETURN;                                 // 提前退出 / Early exit
END_IF
IF (fCloseMin > DL_SEG_HI_MIN) OR (fHeatMin > DL_SEG_HI_MIN)
   OR (fHoldMin > DL_SEG_HI_MIN) OR (fBlowDownMin > DL_SEG_HI_MIN)
   OR (fOpenMin > DL_SEG_HI_MIN) THEN
    fCycleMin := 0.0;                       // 段长越上限：单位多半用错 / Segment too long, unit error likely
    fHoldSharePct := 0.0;                   // 占比不可算 / Share not computable
    xValid := FALSE;                        // 判无效 / Invalid
    FC_DL_TireCureMoldCycleTimeCalc := FALSE;   // 返回码同步 / Return synchronised
    RETURN;                                 // 提前退出 / Early exit
END_IF

(* —— 段 3：主算式（不钳制，先出原始值供段 4 判据使用，R24） —— *)
_fCycleRawMin := fCloseMin + fHeatMin + fHoldMin + fBlowDownMin + fOpenMin;        // 总周期 [min]

(* —— 段 4：总周期零闸（占比式分母） —— *)
IF _fCycleRawMin <= DL_EPS THEN
    fCycleMin := 0.0;                       // 零周期即不可算 / Zero cycle is not computable
    fHoldSharePct := 0.0;                   // 占比不可算 / Share not computable
    xValid := FALSE;                        // 判无效 / Invalid
    FC_DL_TireCureMoldCycleTimeCalc := FALSE;   // 返回码同步 / Return synchronised
    RETURN;                                 // 提前退出 / Early exit
END_IF

_fShareRawPct := fHoldMin / _fCycleRawMin * DL_PCT;                               // 保温段占比 [%]

(* —— 段 5：判据（取原始值；单点 BOOL 聚合避免多处赋 FALSE 覆盖） —— *)
xValid := (_fCycleRawMin <= DL_CYCLE_HI_MIN)                                      // 不超总周期物理上限
          AND (_fShareRawPct >= 0.0)                                              // 占比不得为负
          AND (_fShareRawPct <= DL_PCT_HI);                                       // 占比不得超 100 %

(* —— 段 6：输出单点写盘（钳制到物理域内，判定结果已在段 5 定案） —— *)
fCycleMin := LIMIT(0.0, _fCycleRawMin, DL_CYCLE_HI_MIN);                           // 总周期钳物理域 [min]
fHoldSharePct := LIMIT(0.0, _fShareRawPct, DL_PCT_HI);                             // 占比钳 0..100 [%]
FC_DL_TireCureMoldCycleTimeCalc := xValid;                                         // 返回码：TRUE = 计算可信

END_FUNCTION

(* ---- FC_DL_TireCurePressForceCalc.st ---- *)
(*
  Name: FC_DL_TireCurePressForceCalc
  Category: DL_Process
  Version: 1.0.0
  Round: R91 / 2026-11-25
  开源溯源：clean-room 自研（族 轮胎硫化，ST 开源生态实测 0 命中，无外部代码引入）
  功能：1) 合模力按「胶囊压力 × 轮胎投影面积」计算：
           F = p * A，其中 p 以 kPa 给出、A 以 m2 给出，则
           F[kN] = p[kPa] * 1000[Pa/kPa] * A[m2] / 1000[N/kN] = p * A，
           即数值上 kPa 与 m2 直乘即为 kN，这是本件量纲自证的要点。
        2) 机台额定上限校验：fForceLoadPct = F / fRatedKn * 100，超额定只置 xOverRated 并钳到额定值，
           不把越限值当作可执行指令下发（合模力不足会出明疤，超额定会压伤模具）。
        3) 不足判据：F < fRatedKn * fMinLoadPct / 100 时置 xUnderForce，
           表示胶囊压力不足以撑满花纹（定型不足），供上层提升一次定型压力。
  边界条件：1) 非有限值闸：四路实值入参先过 NOT(x > -DL_BIG AND x < DL_BIG)，同时拦 NaN 与 Inf，
           命中即闸断实值通路（力与负荷率强制 0.0），不得只置标志（R19）。
        2) 面积零闸：轮胎投影面积 fProjectAreaM2 必须 > DL_EPS，否则力恒为零，
           会把「面积未组态」伪装成「无合模力」，因此判无效而非输出 0。
        3) 额定值域闸：fRatedKn 必须 > DL_EPS（负荷率式的分母）；fMinLoadPct 须落在 (0.0, 100.0] 内，
           越域说明阈值未组态（下限为 0 会使不足判据恒假）。
        4) 压力域闸：fPressKpa 不得为负（负表压属传感器错，不取绝对值掩盖）。
        5) 判据取原始值（R24）：超额定与不足判定均使用钳制前的 _fForceRawKn，不得先钳再判。
        6) 物理域钳制：力钳 0.0 ~ fRatedKn；负荷率钳 0.0 ~ DL_PCT_HI。
  量纲自证：p [kPa] = 1000 Pa；A [m2]；p*A = 1000 Pa*m2 = 1000 N = 1 kN，
           故 F[kN] 与 p[kPa]*A[m2] 数值相等，量纲关系合法；
           fForceLoadPct = (kN)/(kN)*100 = 无因次百分数 [%]。
  修订历史 Revision :
    2026-11-25  v1.0.0  R91 首版
*)

FUNCTION FC_DL_TireCurePressForceCalc : BOOL
VAR_INPUT
    fPressKpa        : REAL;   // 胶囊内蒸汽/氮气压力 [kPa] / Bladder steam or nitrogen pressure [kPa]
    fProjectAreaM2   : REAL;   // 轮胎内腔投影面积 [m2] / Tyre inner projection area [m2]
    fRatedKn         : REAL;   // 机台额定合模力 [kN] / Machine rated clamping force [kN]
    fMinLoadPct      : REAL;   // 允许最小负荷率（低于即判定型不足）[%] / Minimum load ratio [%]
END_VAR
VAR_OUTPUT
    fForceKn         : REAL;   // 合模力 [kN] / Clamping force [kN]
    fForceLoadPct    : REAL;   // 合模力对额定值的负荷率 [%] / Load ratio against the rated force [%]
    xUnderForce      : BOOL;   // 合模力不足标志 [bool] / Insufficient clamping force flag [bool]
    xOverRated       : BOOL;   // 超机台额定标志 [bool] / Over rated force flag [bool]
    xValid           : BOOL;   // 计算有效标志 [bool] / Calculation valid flag [bool]
END_VAR
VAR
    _fForceRawKn     : REAL;   // 钳制前的原始合模力 [kN] / Raw clamping force before limiting [kN]
    _fLoadRawPct     : REAL;   // 钳制前的原始负荷率 [%] / Raw load ratio before limiting [%]
    _fMinForceKn     : REAL;   // 允许最小合模力 [kN] / Minimum acceptable clamping force [kN]
END_VAR
VAR CONSTANT
    DL_EPS           : REAL := 1.0E-9;    // 数值零闸阈值 [-] / Numeric zero gate threshold [-]
    DL_BIG           : REAL := 1.0E12;    // 非有限值闸量级上限 [-] / Finiteness gate magnitude [-]
    DL_PCT           : REAL := 100.0;     // 百分比换算因子 [%] / Percent conversion factor [%]
    DL_PCT_HI        : REAL := 100.0;     // 负荷率物理上限 [%] / Load ratio upper bound [%]
END_VAR

(* —— 段 1：非有限值闸（R19：闸断实值通路） —— *)
IF NOT (fPressKpa > -DL_BIG AND fPressKpa < DL_BIG)
   OR NOT (fProjectAreaM2 > -DL_BIG AND fProjectAreaM2 < DL_BIG)
   OR NOT (fRatedKn > -DL_BIG AND fRatedKn < DL_BIG)
   OR NOT (fMinLoadPct > -DL_BIG AND fMinLoadPct < DL_BIG) THEN
    fForceKn := 0.0;                        // 输出强制 0.0，切断污染源 / Force zero, cut polluted path
    fForceLoadPct := 0.0;                   // 负荷率强制 0.0 / Load ratio forced to zero
    xUnderForce := TRUE;                    // 失效侧按不足处理（保守侧）/ Treat as insufficient when invalid
    xOverRated := FALSE;                    // 失效侧超额定位保持假 / Over-rated stays false
    xValid := FALSE;                        // 有效位清零 / Validity cleared
    FC_DL_TireCurePressForceCalc := FALSE;  // 返回码与有效位同源 / Return mirrors validity
    RETURN;                                 // 立即退出 / Immediate exit
END_IF

(* —— 段 2：面积零闸与额定值域闸（面积为乘子，额定值为负荷率分母） —— *)
IF (fProjectAreaM2 <= DL_EPS)                                     // 面积不可为零
   OR (fRatedKn <= DL_EPS)                                        // 额定力必须已组态
   OR (fMinLoadPct <= DL_EPS)                                     // 最小负荷率不可为零（否则判据恒假）
   OR (fMinLoadPct > DL_PCT_HI)                                   // 最小负荷率不得超 100 %
   OR (fPressKpa < 0.0) THEN                                      // 压力不得为负
    fForceKn := 0.0;                        // 参数不可用即无合模力 / No parameter, no force
    fForceLoadPct := 0.0;                   // 负荷率不可算 / Load ratio not computable
    xUnderForce := TRUE;                    // 按不足处理（保守侧）/ Treat as insufficient
    xOverRated := FALSE;                    // 超额定位保持假 / Over-rated stays false
    xValid := FALSE;                        // 判无效 / Invalid
    FC_DL_TireCurePressForceCalc := FALSE;  // 返回码同步 / Return synchronised
    RETURN;                                 // 提前退出 / Early exit
END_IF

(* —— 段 3：主算式（不钳制，先出原始值供段 4 判据使用，R24） —— *)
_fForceRawKn := fPressKpa * fProjectAreaM2;                                       // 合模力 [kN]（kPa*m2 = kN）
_fLoadRawPct := _fForceRawKn / fRatedKn * DL_PCT;                                 // 负荷率 [%]
_fMinForceKn := fRatedKn * fMinLoadPct / DL_PCT;                                  // 允许最小合模力 [kN]

(* —— 段 4：判据（取原始值；单点 BOOL 聚合避免多处赋 FALSE 覆盖） —— *)
xUnderForce := (_fForceRawKn < _fMinForceKn);                                     // 定型不足（压力撑不满花纹）
xOverRated := (_fForceRawKn > fRatedKn);                                          // 超机台额定（压伤模具风险）
xValid := (_fForceRawKn >= 0.0)                                                   // 力不得为负
          AND (_fLoadRawPct >= 0.0)                                               // 负荷率不得为负
          AND (_fMinForceKn >= 0.0);                                              // 最小力不得为负（组态校验）

(* —— 段 5：输出单点写盘（钳制到物理域内，判定结果已在段 4 定案） —— *)
fForceKn := LIMIT(0.0, _fForceRawKn, fRatedKn);                                   // 力钳 0..额定 [kN]
fForceLoadPct := LIMIT(0.0, _fLoadRawPct, DL_PCT_HI);                             // 负荷率钳 0..100 [%]
FC_DL_TireCurePressForceCalc := xValid;                                           // 返回码：TRUE = 计算可信

END_FUNCTION

(* ---- FC_DL_TireCureSteamQualityCalc.st ---- *)
(*
  Name: FC_DL_TireCureSteamQualityCalc
  Category: DL_Process
  Version: 1.0.0
  Round: R91 / 2026-11-25
  开源溯源：clean-room 自研（族 轮胎硫化，ST 开源生态实测 0 命中，无外部代码引入）
  功能：1) 蒸汽干度按焓差法估算：x = (h − h_f) / h_fg，
           h 为实测蒸汽比焓、h_f 为同压力下饱和液比焓、h_fg 为同压力下汽化潜热，
           三者单位一致（kJ/kg），故比值无因次，0 <= x <= 1 即饱和蒸汽的干度区间。
        2) 三态判别（nState）：0 = 饱和蒸汽（0.0 <= x <= 1.0）、1 = 过热蒸汽（x > 1.0）、
           2 = 湿蒸汽/带水（x < 0.0）。硫化工艺要求 x 接近 1.0 的饱和蒸汽，
           带水会显著降低传热系数并在胶囊内壁形成水锤，过热则温度失控。
        3) 干度读数同时钳到 [DL_Q_LO, DL_Q_HI]（-0.5 ~ 1.5），保留三态判别余量，
           避免极端异常值污染趋势曲线。
  边界条件：1) 非有限值闸：三路实值入参先过 NOT(x > -DL_BIG AND x < DL_BIG)，同时拦 NaN 与 Inf，
           命中即闸断实值通路（干度强制 0.0 且 nState 置 2 = 湿蒸汽，保守侧），不得只置标志（R19）。
        2) 分母零闸：汽化潜热 fLatentKjKg 必须 > DL_EPS（干度式分母），否则判无效并清零。
        3) 焓值量级闸：三路焓值必须落在 (0.0, DL_H_HI) 内（水的焓恒为正且不超过 4000 kJ/kg 量级），
           越域说明单位用错（J 与 kJ 混用）或测点失效，判无效。
        4) 一致性校验：h_f + h_fg 必须与 h 同量级 —— 若 h_f + h_fg <= DL_EPS，说明压力对应的
           饱和参数未组态（表查错），判无效而非硬算。
        5) 判据取原始值（R24）：三态判别使用钳制前的 _fQualityRaw，不得先钳再判。
        6) 纯函数无状态：干度的滑动平均与趋势判断由上层蒸汽品质监视模块承担。
  量纲自证：x = (kJ/kg − kJ/kg) / (kJ/kg) = 无因次 [-]，量纲合法；
           nState 为无量纲枚举等级 [level]。
  修订历史 Revision :
    2026-11-25  v1.0.0  R91 首版
*)

FUNCTION FC_DL_TireCureSteamQualityCalc : BOOL
VAR_INPUT
    fEnthalpyKjKg    : REAL;   // 实测蒸汽比焓 [kJ/kg] / Measured steam specific enthalpy [kJ/kg]
    fSatLiqEnthKjKg  : REAL;   // 同压力下饱和液比焓 [kJ/kg] / Saturated liquid enthalpy at the same pressure [kJ/kg]
    fLatentKjKg      : REAL;   // 同压力下汽化潜热 [kJ/kg] / Latent heat of vaporisation at the same pressure [kJ/kg]
END_VAR
VAR_OUTPUT
    fQuality         : REAL;   // 蒸汽干度（无因次）[-] / Steam quality, dimensionless [-]
    nState           : INT;    // 三态判别 0=饱和 1=过热 2=湿蒸汽/带水 [level] / Steam state 0/1/2 [level]
    xValid           : BOOL;   // 计算有效标志 [bool] / Calculation valid flag [bool]
END_VAR
VAR
    _fQualityRaw     : REAL;   // 钳制前的原始干度 [-]/ Raw quality before limiting [-]
END_VAR
VAR CONSTANT
    DL_EPS           : REAL := 1.0E-9;    // 数值零闸阈值 [-] / Numeric zero gate threshold [-]
    DL_BIG           : REAL := 1.0E12;    // 非有限值闸量级上限 [-] / Finiteness gate magnitude [-]
    DL_H_HI          : REAL := 4000.0;    // 焓值量级上限 [kJ/kg] / Enthalpy magnitude upper bound [kJ/kg]
    DL_Q_LO          : REAL := -0.5;      // 干度显示下限 [-]/ Quality display low bound [-]
    DL_Q_HI          : REAL := 1.5;       // 干度显示上限 [-]/ Quality display high bound [-]
    DL_Q_SAT_HI      : REAL := 1.0;       // 饱和蒸汽干度上限 [-]/ Saturated steam quality upper bound [-]
    DL_ST_SAT        : INT := 0;          // 三态：饱和蒸汽 [level] / State: saturated steam [level]
    DL_ST_SUPER      : INT := 1;          // 三态：过热蒸汽 [level] / State: superheated steam [level]
    DL_ST_WET        : INT := 2;          // 三态：湿蒸汽/带水 [level] / State: wet steam with water [level]
END_VAR

(* —— 段 1：非有限值闸（R19：闸断实值通路；失效侧置湿蒸汽，保守侧） —— *)
IF NOT (fEnthalpyKjKg > -DL_BIG AND fEnthalpyKjKg < DL_BIG)
   OR NOT (fSatLiqEnthKjKg > -DL_BIG AND fSatLiqEnthKjKg < DL_BIG)
   OR NOT (fLatentKjKg > -DL_BIG AND fLatentKjKg < DL_BIG) THEN
    fQuality := 0.0;                        // 输出强制 0.0，切断污染源 / Force zero, cut polluted path
    nState := DL_ST_WET;                    // 失效侧按带水处理（保守侧：宁可拒用不可误用）
    xValid := FALSE;                        // 有效位清零 / Validity cleared
    FC_DL_TireCureSteamQualityCalc := FALSE;   // 返回码与有效位同源 / Return mirrors validity
    RETURN;                                 // 立即退出 / Immediate exit
END_IF

(* —— 段 2：分母零闸（潜热为干度式分母） —— *)
IF fLatentKjKg <= DL_EPS THEN
    fQuality := 0.0;                        // 潜热缺失即不可算 / No latent heat, no quality
    nState := DL_ST_WET;                    // 按带水处理（保守侧）/ Treat as wet steam
    xValid := FALSE;                        // 判无效 / Invalid
    FC_DL_TireCureSteamQualityCalc := FALSE;   // 返回码同步 / Return synchronised
    RETURN;                                 // 提前退出 / Early exit
END_IF

(* —— 段 3：焓值量级闸与饱和参数一致性闸（防单位混用与测点失效） —— *)
IF (fEnthalpyKjKg <= 0.0) OR (fEnthalpyKjKg >= DL_H_HI)
   OR (fSatLiqEnthKjKg < 0.0) OR (fSatLiqEnthKjKg >= DL_H_HI)
   OR (fLatentKjKg >= DL_H_HI)
   OR ((fSatLiqEnthKjKg + fLatentKjKg) <= DL_EPS) THEN
    fQuality := 0.0;                        // 焓值越域即不可算 / Enthalpy out of range
    nState := DL_ST_WET;                    // 按带水处理（保守侧）/ Treat as wet steam
    xValid := FALSE;                        // 判无效 / Invalid
    FC_DL_TireCureSteamQualityCalc := FALSE;   // 返回码同步 / Return synchronised
    RETURN;                                 // 提前退出 / Early exit
END_IF

(* —— 段 4：主算式（不钳制，先出原始值供段 5 判据使用，R24） —— *)
_fQualityRaw := (fEnthalpyKjKg - fSatLiqEnthKjKg) / fLatentKjKg;                  // 干度 [-]

(* —— 段 5：三态判别（取原始值；判别顺序由湿到过，互斥且完整） —— *)
IF _fQualityRaw < 0.0 THEN
    nState := DL_ST_WET;                    // 带水
ELSIF _fQualityRaw > DL_Q_SAT_HI THEN
    nState := DL_ST_SUPER;                  // 过热
ELSE
    nState := DL_ST_SAT;                    // 饱和
END_IF

xValid := (_fQualityRaw >= DL_Q_LO)                                               // 低于显示下限属量级异常
          AND (_fQualityRaw <= DL_Q_HI);                                          // 高于显示上限属量级异常

(* —— 段 6：输出单点写盘（钳制到显示域内，判别结果已在段 5 定案） —— *)
fQuality := LIMIT(DL_Q_LO, _fQualityRaw, DL_Q_HI);                                // 干度钳 -0.5..1.5 [-]
FC_DL_TireCureSteamQualityCalc := xValid;                                         // 返回码：TRUE = 计算可信

END_FUNCTION

(* ---- FC_DL_TireCureTempGradientCalc.st ---- *)
(*
  Name: FC_DL_TireCureTempGradientCalc
  Category: DL_Process
  Version: 1.0.0
  Round: R91 / 2026-11-25
  开源溯源：clean-room 自研（族 轮胎硫化，ST 开源生态实测 0 命中，无外部代码引入）
  功能：1) 胎面温差按「外表面温度与内表面温度之差」计算：dT = T_outer − T_inner；
           方向固定不可交换（热流由外模经胎体传向内腔），负值表示测温点接反。
        2) 温度梯度按温差除以导热路径长度折算：grad = dT / (path_mm / 1000)，单位 K/m，
           用于判断硫化过程中胎体内部是否处于「急热」状态（梯度大易产生内部应力与海绵）。
           同时给出以 K/mm 计的分级量 fGradKmm，方便工艺按毫米壁厚直观比对。
        3) 温差超限分级（nGrade）：0 = 正常（dT <= fDeltaWarnK）、1 = 预警（<= fDeltaMaxK）、
           2 = 超限（> fDeltaMaxK），供上层决定是否延长预热段或降低外模温度。
  边界条件：1) 非有限值闸：五路实值入参先过 NOT(x > -DL_BIG AND x < DL_BIG)，同时拦 NaN 与 Inf，
           命中即闸断实值通路（温差与梯度强制 0.0 且分级置 2 = 超限），不得只置标志（R19）。
        2) 路径零闸：导热路径 fPathMm 必须 > DL_EPS（梯度的分母），否则判无效并清零。
        3) 分级阈值域闸：须满足 0.0 < fDeltaWarnK < fDeltaMaxK，否则两级判据区间为空、分级恒失效，
           越域判无效并把 nGrade 置 2（保守侧）。
        4) 温差方向闸：dT 必须 > 0（外表面必须比内表面热），为负属测点错位，判无效，
           不取绝对值掩盖符号错误。
        5) 判据取原始值（R24）：分级使用原始温差与原始梯度，钳制只作用于输出数值。
        6) 物理域钳制：温差钳 0.0 ~ DL_DELTA_HI；梯度钳 0.0 ~ DL_GRAD_HI。
  量纲自证：dT = (degC) − (degC) = (K)；
           grad = (K)/(m) = K/m，另 (K)/(mm) = K/mm；
           两条梯度量同源于 dT 与 path，属同一量纲族的不同长度基准，均已显式标注。
  修订历史 Revision :
    2026-11-25  v1.0.0  R91 首版
*)

FUNCTION FC_DL_TireCureTempGradientCalc : BOOL
VAR_INPUT
    fOuterC          : REAL;   // 胎面外表面温度 [degC] / Tread outer surface temperature [degC]
    fInnerC          : REAL;   // 胎体内表面温度 [degC] / Tyre inner surface temperature [degC]
    fPathMm          : REAL;   // 外表面到内表面的导热路径长度 [mm] / Conduction path length [mm]
    fDeltaWarnK      : REAL;   // 温差预警阈值 [K] / Temperature difference warning threshold [K]
    fDeltaMaxK       : REAL;   // 温差上限阈值 [K] / Temperature difference upper limit [K]
END_VAR
VAR_OUTPUT
    fDeltaTK         : REAL;   // 胎面温差 [K] / Tread temperature difference [K]
    fGradKmm         : REAL;   // 以毫米为基准的温度梯度 [K/mm] / Gradient per millimetre [K/mm]
    fGradKm          : REAL;   // 以米为基准的温度梯度 [K/m] / Gradient per metre [K/m]
    nGrade           : INT;    // 温差分级 0=正常 1=预警 2=超限 [level] / Difference grade 0/1/2 [level]
    xValid           : BOOL;   // 计算有效标志 [bool] / Calculation valid flag [bool]
END_VAR
VAR
    _fDeltaRawK      : REAL;   // 钳制前的原始温差 [K] / Raw temperature difference [K]
    _fGradRawKmm     : REAL;   // 钳制前的原始梯度 [K/mm] / Raw gradient before limiting [K/mm]
    _fGradRawKm      : REAL;   // 钳制前的原始梯度 [K/m] / Raw gradient per metre [K/m]
END_VAR
VAR CONSTANT
    DL_EPS           : REAL := 1.0E-9;    // 数值零闸阈值 [-] / Numeric zero gate threshold [-]
    DL_BIG           : REAL := 1.0E12;    // 非有限值闸量级上限 [-] / Finiteness gate magnitude [-]
    DL_MM_PER_M      : REAL := 1000.0;    // 米到毫米的折算 [mm/m] / Millimetres per metre [mm/m]
    DL_DELTA_HI      : REAL := 500.0;     // 温差物理上限 [K] / Temperature difference upper bound [K]
    DL_GRAD_HI       : REAL := 1000.0;    // 梯度物理上限 [K/m] / Gradient upper bound [K/m]
    DL_GRADE_OK      : INT := 0;          // 分级：正常 [level] / Grade: normal [level]
    DL_GRADE_WARN    : INT := 1;          // 分级：预警 [level] / Grade: warning [level]
    DL_GRADE_BAD     : INT := 2;          // 分级：超限 [level] / Grade: out of limit [level]
END_VAR

(* —— 段 1：非有限值闸（R19：闸断实值通路；失效侧分级置超限） —— *)
IF NOT (fOuterC > -DL_BIG AND fOuterC < DL_BIG)
   OR NOT (fInnerC > -DL_BIG AND fInnerC < DL_BIG)
   OR NOT (fPathMm > -DL_BIG AND fPathMm < DL_BIG)
   OR NOT (fDeltaWarnK > -DL_BIG AND fDeltaWarnK < DL_BIG)
   OR NOT (fDeltaMaxK > -DL_BIG AND fDeltaMaxK < DL_BIG) THEN
    fDeltaTK := 0.0;                        // 输出强制 0.0，切断污染源 / Force zero, cut polluted path
    fGradKmm := 0.0;                        // 梯度强制 0.0 / Gradient forced to zero
    fGradKm := 0.0;                         // 梯度强制 0.0 / Gradient forced to zero
    nGrade := DL_GRADE_BAD;                 // 失效侧按超限处理（保守侧）/ Treat as out of limit when invalid
    xValid := FALSE;                        // 有效位清零 / Validity cleared
    FC_DL_TireCureTempGradientCalc := FALSE;   // 返回码与有效位同源 / Return mirrors validity
    RETURN;                                 // 立即退出 / Immediate exit
END_IF

(* —— 段 2：路径零闸与阈值域闸 —— *)
IF (fPathMm <= DL_EPS)                                            // 路径不可为零（梯度分母）
   OR (fDeltaWarnK <= DL_EPS)                                     // 预警阈值必须为正
   OR (fDeltaMaxK <= fDeltaWarnK) THEN                            // 上限必须严格大于预警阈值
    fDeltaTK := 0.0;                        // 参数不可用即无温差 / No parameter, no difference
    fGradKmm := 0.0;                        // 梯度不可算 / Gradient not computable
    fGradKm := 0.0;                         // 梯度不可算 / Gradient not computable
    nGrade := DL_GRADE_BAD;                 // 按超限处理（保守侧）/ Treat as out of limit
    xValid := FALSE;                        // 判无效 / Invalid
    FC_DL_TireCureTempGradientCalc := FALSE;   // 返回码同步 / Return synchronised
    RETURN;                                 // 提前退出 / Early exit
END_IF

(* —— 段 3：主算式（不钳制，先出原始值供段 4 判据使用，R24） —— *)
_fDeltaRawK := fOuterC - fInnerC;                                                 // 胎面温差 [K]
_fGradRawKmm := _fDeltaRawK / fPathMm;                                            // 梯度 [K/mm]
_fGradRawKm := _fDeltaRawK / (fPathMm / DL_MM_PER_M);                             // 梯度 [K/m]

(* —— 段 4：判据与分级（取原始值；单点 BOOL 聚合避免多处赋 FALSE 覆盖） —— *)
xValid := (_fDeltaRawK > 0.0)                                                     // 外表面必须比内表面热（方向固定）
          AND (_fDeltaRawK <= DL_DELTA_HI)                                        // 不超温差物理上限
          AND (_fGradRawKm > 0.0)                                                 // 梯度必须为正
          AND (_fGradRawKm <= DL_GRAD_HI)                                         // 不超梯度物理上限
          AND (fDeltaMaxK <= DL_DELTA_HI);                                        // 上限阈值须在物理域内

IF NOT xValid THEN
    nGrade := DL_GRADE_BAD;                 // 参数非法：按超限处理（保守侧）
ELSIF _fDeltaRawK > fDeltaMaxK THEN
    nGrade := DL_GRADE_BAD;                 // 温差超上限
ELSIF _fDeltaRawK > fDeltaWarnK THEN
    nGrade := DL_GRADE_WARN;                // 预警带
ELSE
    nGrade := DL_GRADE_OK;                  // 正常
END_IF

(* —— 段 5：输出单点写盘（钳制到物理域内，分级已在段 4 定案） —— *)
fDeltaTK := LIMIT(0.0, _fDeltaRawK, DL_DELTA_HI);                                  // 温差钳物理域 [K]
fGradKmm := LIMIT(0.0, _fGradRawKmm, DL_GRAD_HI);                                  // 梯度钳物理域 [K/mm]
fGradKm := LIMIT(0.0, _fGradRawKm, DL_GRAD_HI);                                    // 梯度钳物理域 [K/m]
FC_DL_TireCureTempGradientCalc := xValid;                                         // 返回码：TRUE = 计算可信

END_FUNCTION

(* ---- FC_DL_TobaccoComponentRatioCalc.st ---- *)
(*
 * FC_DL_TobaccoComponentRatioCalc | C1 | DL_Process
 * 功能：叶丝/梗丝/膨胀丝三组分掺配比例求和、平衡判定与主组分识别       单位：比例 [%]、主组分为序号 1/2/3
 * 工况边界：三比例须均为有限且 ≥0；任一为负即判 9501 并置 xValid=FALSE（所有出口取安全值）；平衡判据为 Σ=100±0.1 %，浮点比较用容差而非相等
 * 代数值回代：70.0 / 20.0 / 10.0 → Σ=100.0、|Σ−100|=0 ≤0.1 → xBalanced=TRUE、nDominant=1（叶丝）
 * 开源溯源：clean-room 自研，未复制任何第三方代码（无外部来源）
 *)
FUNCTION FC_DL_TobaccoComponentRatioCalc : BOOL
VAR_INPUT
    rLeafCutPct  : REAL;             // 叶丝比例 | leaf cut tobacco ratio [%]
    rStemCutPct  : REAL;             // 梗丝比例 | stem cut tobacco ratio [%]
    rExpandedPct : REAL;             // 膨胀丝比例 | expanded tobacco ratio [%]
END_VAR
VAR_OUTPUT
    rSumPct     : REAL;              // 三组分之和 | sum of the three components [%]
    xBalanced   : BOOL;              // 配比平衡（Σ=100±0.1）| ratio balanced within 100 ± 0.1 [%]
    nDominant   : INT;               // 主组分：1=叶丝 / 2=梗丝 / 3=膨胀丝 | dominant component index
    xValid      : BOOL;              // 输出有效 | outputs valid
    nFaultCode  : INT;               // 0=无 / 9501=组分比例非法 | 0 none, 9501 illegal component ratio
END_VAR
VAR
    xFinA : BOOL;                    // 叶丝比例有限性 | leaf ratio is finite
    xFinB : BOOL;                    // 梗丝比例有限性 | stem ratio is finite
    xFinC : BOOL;                    // 膨胀丝比例有限性 | expanded ratio is finite
END_VAR
VAR CONSTANT
    DL_TCR_TOTAL : REAL := 100.0;    // 配比总和基准 | total ratio reference [%]
    DL_TCR_TOL   : REAL := 0.1;      // 平衡容差 | balance tolerance [%]
    DL_TCR_EPS   : REAL := 1.0E-6;   // 浮点比较容差 | floating comparison tolerance [%]
END_VAR

// 段1｜非有限闸（R19）
xFinA := (rLeafCutPct = rLeafCutPct) AND ((rLeafCutPct - rLeafCutPct) = 0.0);
xFinB := (rStemCutPct = rStemCutPct) AND ((rStemCutPct - rStemCutPct) = 0.0);
xFinC := (rExpandedPct = rExpandedPct) AND ((rExpandedPct - rExpandedPct) = 0.0);
IF (NOT xFinA) OR (NOT xFinB) OR (NOT xFinC) THEN
    rSumPct := 0.0;                  // 安全值：和 0 | safe value, zero sum
    xBalanced := FALSE;
    nDominant := 0;
    xValid := FALSE;
    nFaultCode := 9501;
    FC_DL_TobaccoComponentRatioCalc := FALSE;
    RETURN;
END_IF

// 段2｜域闸：任一比例为负即判非法
IF (rLeafCutPct < 0.0) OR (rStemCutPct < 0.0) OR (rExpandedPct < 0.0) THEN
    rSumPct := 0.0;
    xBalanced := FALSE;
    nDominant := 0;
    xValid := FALSE;
    nFaultCode := 9501;
    FC_DL_TobaccoComponentRatioCalc := FALSE;
    RETURN;
END_IF

// 段3｜求和与平衡判定
rSumPct := rLeafCutPct + rStemCutPct + rExpandedPct;
xBalanced := ABS(rSumPct - DL_TCR_TOTAL) <= (DL_TCR_TOL + DL_TCR_EPS);

// 段4｜主组分识别（严格大于，等值时按叶丝优先，避免不确定主组分）
nDominant := 1;
IF (rStemCutPct > rLeafCutPct) AND (rStemCutPct >= rExpandedPct) THEN
    nDominant := 2;
ELSIF (rExpandedPct > rLeafCutPct) AND (rExpandedPct > rStemCutPct) THEN
    nDominant := 3;
END_IF

// 段5｜出口
nFaultCode := 0;
xValid := TRUE;
FC_DL_TobaccoComponentRatioCalc := TRUE;
END_FUNCTION

(* ---- FC_DL_TobaccoFillValueCalc.st ---- *)
(*
 * FC_DL_TobaccoFillValueCalc | C1 | DL_Process
 * 功能：烟丝填充值（松装单位质量体积）与工艺区间判定       单位：质量 [g]、体积 [mL]，填充值 [cm³/g]
 * 工况边界：仅适用于松装法（标准量筒自由落料）测量；样品质量须 >0（入分母）；膨胀丝填充值工艺区间 8~12 cm³/g，超出仅置信息位不判故障
 * 代数值回代：m=50 g、V=500 mL → FV=500/50=10.0 cm³/g，落在 8~12 → xInRange=TRUE（与 spec 回代行一致）
 * 开源溯源：clean-room 自研，未复制任何第三方代码（无外部来源）
 *)
FUNCTION FC_DL_TobaccoFillValueCalc : BOOL
VAR_INPUT
    rSampleMassG    : REAL := 50.0;   // 样品质量 | sample mass [g]
    rCylinderVolMl  : REAL := 500.0;  // 量筒松装体积 | loose bulk volume in the cylinder [mL]
END_VAR
VAR_OUTPUT
    rFillValueCm3g : REAL;            // 填充值 | fill value [cm³/g]
    xInRange       : BOOL;            // 落在膨胀丝工艺区间 8~12 | inside the expanded tobacco range 8 to 12
    xValid         : BOOL;            // 输出有效 | outputs valid
    nFaultCode     : INT;             // 0=无 / 9511=样品质量或体积非法 | 0 none, 9511 illegal sample mass or volume
END_VAR
VAR
    xFinMass : BOOL;                  // 质量有限性 | mass is finite
    xFinVol  : BOOL;                  // 体积有限性 | volume is finite
END_VAR
VAR CONSTANT
    DL_TFV_MASS_MIN : REAL := 1.0E-6;  // 质量下限（防零除）| mass lower bound guarding the division [g]
    DL_TFV_RANGE_LO : REAL := 8.0;     // 工艺区间下限 | process range lower bound [cm³/g]
    DL_TFV_RANGE_HI : REAL := 12.0;    // 工艺区间上限 | process range upper bound [cm³/g]
    DL_TFV_EPS      : REAL := 1.0E-6;  // 浮点比较容差 | floating comparison tolerance [cm³/g]
END_VAR

// 段1｜非有限闸（R19）
xFinMass := (rSampleMassG = rSampleMassG) AND ((rSampleMassG - rSampleMassG) = 0.0);
xFinVol := (rCylinderVolMl = rCylinderVolMl) AND ((rCylinderVolMl - rCylinderVolMl) = 0.0);
IF (NOT xFinMass) OR (NOT xFinVol) THEN
    rFillValueCm3g := 0.0;            // 安全值：填充值 0 | safe value, zero fill value
    xInRange := FALSE;
    xValid := FALSE;
    nFaultCode := 9511;
    FC_DL_TobaccoFillValueCalc := FALSE;
    RETURN;
END_IF

// 段2｜域闸：质量入分母必须 >0，体积必须 >0
IF (rSampleMassG <= DL_TFV_MASS_MIN) OR (rCylinderVolMl <= 0.0) THEN
    rFillValueCm3g := 0.0;
    xInRange := FALSE;
    xValid := FALSE;
    nFaultCode := 9511;
    FC_DL_TobaccoFillValueCalc := FALSE;
    RETURN;
END_IF

// 段3｜算法：FV = V/m（mL = cm³，量纲直接相通）
rFillValueCm3g := rCylinderVolMl / rSampleMassG;

// 段4｜区间判定（判据与出口同源于原始测量值）
xInRange := (rFillValueCm3g >= (DL_TFV_RANGE_LO - DL_TFV_EPS))
             AND (rFillValueCm3g <= (DL_TFV_RANGE_HI + DL_TFV_EPS));
nFaultCode := 0;
xValid := TRUE;
FC_DL_TobaccoFillValueCalc := TRUE;
END_FUNCTION

(* ---- FC_DL_UnderflowDensityCalc.st ---- *)
(*
  Name: FC_DL_UnderflowDensityCalc
  Category: DL_Process
  Version: 1.0.0
  Round: R89 / 2026-11-25
  开源溯源：clean-room 自研（族 矿山破碎筛分，ST 开源生态实测 0 命中，无外部代码引入）
  功能：由底流管压力变送器读数与取压点高度反算浆体密度，再换算底流固体质量浓度与体积浓度。
  边界条件：① 四入参全部过非有限闸，任一非有限返回哨兵 -1；
            ② 取压点高度为除子（P = ρ·g·h 反解），须 0.2~20 m；压力须 ≥ 0 且 ≤ 500 kPa；
            ③ 固体密度必须高于浆体密度且高于水密度，否则质量浓度式分母塌零或无物理意义，返回哨兵 -1；
            ④ 质量浓度物理域 0~100 %，越域（传感器零漂）判非法返回哨兵 -1，不静默钳位。
  量纲自证：P[kPa]×1000 = Pa = N/m2；N/m2 ÷ (m/s2 × m) = kg/m3；浓度式无量纲。
*)
FUNCTION FC_DL_UnderflowDensityCalc : REAL
VAR_INPUT
    fPressKPa : REAL;            (* 取压点表压 [kPa] Gauge pressure at tapping point [kPa] *)
    fHeightM : REAL;             (* 取压点距液面高度 [m] Tapping height below surface [m] *)
    fSlurryDensityKgM3 : REAL;   (* 浆体密度（用于浓度换算的复核值） [kg/m3] Slurry density [kg/m3] *)
    fSolidDensityKgM3 : REAL;    (* 固体真密度 [kg/m3] Solids true density [kg/m3] *)
END_VAR
VAR_OUTPUT
    fMassConcPct : REAL;         (* 固体质量浓度 [%] Solids mass concentration [%] *)
    fVolConcPct : REAL;          (* 固体体积浓度 [%] Solids volume concentration [%] *)
    xValid : BOOL;               (* 计算有效性标志 [-] Calculation valid flag *)
END_VAR
VAR CONSTANT
    DL_EPS : REAL := 1.0E-9;         (* 除零判定容差 [-] Divide-by-zero tolerance *)
    DL_G : REAL := 9.80665;          (* 标准重力加速度 [m/s2] Standard gravity [m/s2] *)
    DL_RHO_W : REAL := 998.2;        (* 水密度（20 ℃） [kg/m3] Water density at 20 degC [kg/m3] *)
    DL_PCT : REAL := 100.0;          (* 百分数基准 [%] Percent base *)
    DL_PA_PER_KPA : REAL := 1000.0;  (* kPa → Pa 换算 [Pa/kPa] Kilopascal to pascal *)
    DL_H_MIN : REAL := 0.2;          (* 取压高度下限 [m] Tapping height floor [m] *)
    DL_H_MAX : REAL := 20.0;         (* 取压高度上限 [m] Tapping height ceiling [m] *)
    DL_P_MAX : REAL := 500.0;        (* 压力上限 [kPa] Pressure ceiling [kPa] *)
    DL_SL_MIN : REAL := 1000.0;      (* 浆体密度下限 [kg/m3] Slurry density floor [kg/m3] *)
    DL_SL_MAX : REAL := 2200.0;      (* 浆体密度上限 [kg/m3] Slurry density ceiling [kg/m3] *)
    DL_SD_MIN : REAL := 1500.0;      (* 固体密度下限 [kg/m3] Solids density floor [kg/m3] *)
    DL_SD_MAX : REAL := 5000.0;      (* 固体密度上限 [kg/m3] Solids density ceiling [kg/m3] *)
END_VAR
VAR
    fRhoCalc : REAL;    (* 由压差反算的浆体密度 [kg/m3] Slurry density from pressure [kg/m3] *)
    fDensDiff : REAL;   (* 固液密度差 [kg/m3] Solids minus water density [kg/m3] *)
    fCm : REAL;         (* 质量浓度小数 [-] Mass concentration fraction *)
END_VAR
(* 出口预置：三出口统一预置（R256） *)
fMassConcPct := 0.0; fVolConcPct := 0.0; xValid := FALSE;
(* 非有限闸：NaN 自反判 + Inf 差值自减判，四入参全枚举 *)
IF (fPressKPa <> fPressKPa) OR ((fPressKPa - fPressKPa) <> 0.0)
   OR (fHeightM <> fHeightM) OR ((fHeightM - fHeightM) <> 0.0)
   OR (fSlurryDensityKgM3 <> fSlurryDensityKgM3) OR ((fSlurryDensityKgM3 - fSlurryDensityKgM3) <> 0.0)
   OR (fSolidDensityKgM3 <> fSolidDensityKgM3) OR ((fSolidDensityKgM3 - fSolidDensityKgM3) <> 0.0) THEN
    FC_DL_UnderflowDensityCalc := -1.0;     (* 哨兵 -1：入参非有限 / Sentinel -1, non-finite input *)
    RETURN;
END_IF
(* 组态域闸：高度为除子，两密度须物理可行且固相明显重于液相 *)
IF (fHeightM < DL_H_MIN) OR (fHeightM > DL_H_MAX)
   OR (fPressKPa < 0.0) OR (fPressKPa > DL_P_MAX)
   OR (fSlurryDensityKgM3 < DL_SL_MIN) OR (fSlurryDensityKgM3 > DL_SL_MAX)
   OR (fSolidDensityKgM3 < DL_SD_MIN) OR (fSolidDensityKgM3 > DL_SD_MAX)
   OR ((fSolidDensityKgM3 - fSlurryDensityKgM3) < DL_EPS) THEN
    FC_DL_UnderflowDensityCalc := -1.0;     (* 哨兵 -1：组态非法 / Sentinel -1, bad configuration *)
    RETURN;
END_IF
(* 反算浆体密度：ρ = P/(g·h)，量纲 Pa ÷ (m/s2·m) = kg/m3 *)
fRhoCalc := (fPressKPa * DL_PA_PER_KPA) / (DL_G * fHeightM);
(* 固液密度差已过正性闸，绝无零除 *)
fDensDiff := fSolidDensityKgM3 - DL_RHO_W;
(* 质量浓度：Cm = ρs(ρsl − ρw) / (ρsl(ρs − ρw))，无量纲 *)
IF fRhoCalc <= DL_EPS THEN
    FC_DL_UnderflowDensityCalc := -1.0;     (* 哨兵 -1：反算密度塌零 / Sentinel -1, vanishing density *)
    RETURN;
END_IF
fCm := (fSolidDensityKgM3 * (fRhoCalc - DL_RHO_W)) / (fRhoCalc * fDensDiff);
(* 物理域检查：质量浓度越 0~1 说明零漂或密度参数不匹配，判非法不钳位 *)
IF (fCm < 0.0) OR (fCm > 1.0) THEN
    FC_DL_UnderflowDensityCalc := -1.0;     (* 哨兵 -1：浓度越物理域 / Sentinel -1, out of physical domain *)
    RETURN;
END_IF
fMassConcPct := fCm * DL_PCT;
(* 体积浓度：Cv = Cm·ρsl/ρs *)
fVolConcPct := (fCm * fRhoCalc / fSolidDensityKgM3) * DL_PCT;
xValid := TRUE;                             (* 链路有效 / Chain valid *)
FC_DL_UnderflowDensityCalc := fMassConcPct;
END_FUNCTION

(* ---- FC_DL_VenturiScrubDpEst.st ---- *)
(*
  道莅工业代码库 / Daoli Industrial ST Library
  组件: FC_DL_VenturiScrubDpEst
  分类: DL_Process
  开源溯源: 无（clean-room 工程公式自研；参考公开工艺计算公式，未复制任何受版权保护代码）
  许可证: 本项目自有 (MIT)
  功能: 文丘里洗涤器喉口压降估算（干气流速头 × 液气动量耦合系数）
  简化式声明: ΔP[kPa] = (ρg·v²/2)·(1 + 0.10·(L/Q)[L每m3]) / 1000；
              0.10 为厂商公开资料常用的液气动量耦合经验系数，非热力学严格值
*)
FUNCTION FC_DL_VenturiScrubDpEst : BOOL
VAR_INPUT
    rGasM3h : REAL; // 实际工况烟气量 [m3/h] / actual gas flow
    rThroatDm : REAL; // 喉口直径 [dm] / throat diameter in decimetre
    rLiquidLM3h : REAL; // 喷液量 [L/h] / sprayed liquid flow
    rRhoGas : REAL; // 工况气体密度 [kg/m3] / gas density at working conditions
END_VAR
VAR_OUTPUT
    rDpKpa : REAL; // 喉口压降 [kPa] / throat pressure drop
    bValid : BOOL; // 结果有效位 [-] / result valid flag
    iErrCode : INT; // 事件码 0=正常 1=喉口直径非法 2=烟气量非法 3=气体密度非法 4=结果非有限 / event code
END_VAR
VAR CONSTANT
    rPi : REAL := 3.14159265358979; // 圆周率 [-] / pi
    rDmToM : REAL := 0.1; // 分米转米系数 [m/dm] / decimetre to metre factor
    rSecPerHour : REAL := 3600.0; // 每小时秒数 [s/h] / seconds per hour
    rPaToKpa : REAL := 0.001; // 帕转千帕系数 [kPa/Pa] / pascal to kilopascal factor
    rLgCoef : REAL := 0.10; // 液气动量耦合经验系数 [-] / empirical liquid-gas momentum coefficient
    rM3ToL : REAL := 1000.0; // 立方米转升系数 [L/m3] / cubic metre to litre factor
END_VAR
VAR
    rDmM : REAL; // 喉口直径 [m] / throat diameter in metre
    rAreaM2 : REAL; // 喉口截面积 [m2] / throat area
    rVelMs : REAL; // 喉口气速 [m/s] / throat gas velocity
    rLgRatio : REAL; // 液气比 [L/m3] / liquid to gas ratio
    rDpPa : REAL; // 压降 [Pa] / pressure drop in pascal
END_VAR

    // —— 段 0：全路径预清 —— //
    rDmM := 0.0;
    rAreaM2 := 0.0;
    rVelMs := 0.0;
    rLgRatio := 0.0;
    rDpPa := 0.0;
    rDpKpa := 0.0;
    bValid := FALSE;
    iErrCode := 0;
    FC_DL_VenturiScrubDpEst := FALSE;
    // —— 段 1：分母闸（喉口直径、烟气量）与密度域闸 —— //
    IF rThroatDm <= 0.0 THEN
        iErrCode := 1; // 喉口直径非法，截面积无定义 / invalid throat diameter
        RETURN;
    END_IF;
    IF rGasM3h <= 0.0 THEN
        iErrCode := 2; // 烟气量非法，气速无定义 / invalid gas flow, velocity undefined
        RETURN;
    END_IF;
    IF rRhoGas <= 0.0 THEN
        iErrCode := 3; // 气体密度非法 / invalid gas density
        RETURN;
    END_IF;
    // —— 段 2：喉口几何与气速（量纲 (m3/h)/(s/h)/(m2) = m/s） —— //
    rDmM := rThroatDm * rDmToM; // 喉口直径 [m] / throat diameter
    rAreaM2 := rPi * rDmM * rDmM / 4.0; // 喉口面积 [m2] / throat area
    IF rAreaM2 <= 1.0E-9 THEN
        iErrCode := 1; // 面积退化，视为直径非法 / degenerate area, treat as invalid diameter
        RETURN;
    END_IF;
    rVelMs := rGasM3h / rSecPerHour / rAreaM2; // 喉口气速 [m/s] / throat velocity
    rLgRatio := rLiquidLM3h / rGasM3h * rM3ToL; // 液气比 [L/m3] / liquid to gas ratio
    // —— 段 3：压降估算（量纲 (kg/m3)*(m2/s2) = Pa） —— //
    rDpPa := (rRhoGas * rVelMs * rVelMs / 2.0) * (1.0 + rLgCoef * rLgRatio); // 压降 [Pa] / pressure drop
    IF ABS(rDpPa) > 1.0E15 THEN
        iErrCode := 4; // 结果非有限，强制归零 / non-finite result, forced to zero
        RETURN;
    END_IF;
    // —— 段 4：单位换算与负值防御 —— //
    IF rDpPa < 0.0 THEN
        rDpKpa := 0.0; // 负输入防御 / negative input guard
    ELSE
        rDpKpa := rDpPa * rPaToKpa; // 压降 [kPa] / pressure drop in kPa
    END_IF;
    bValid := TRUE;
    FC_DL_VenturiScrubDpEst := TRUE;
END_FUNCTION

(* ---- FC_DL_VfaAlkalinityRatio.st ---- *)
(*
  道莅工业代码库 / Daoli Industrial ST Library
  组件: FC_DL_VfaAlkalinityRatio
  分类: DL_Process
  开源溯源: 无（clean-room 工程公式自研；参考公开工艺计算公式，未复制任何受版权保护代码）
  许可证: 本项目自有 (MIT)
  功能: VFA/碱度比计算与酸化风险分级（0=正常 1=关注 2=酸化预警）
*)
FUNCTION FC_DL_VfaAlkalinityRatio : BOOL
VAR_INPUT
    rVfaMgL : REAL; // 挥发性脂肪酸浓度 [mg/L，以乙酸计] / volatile fatty acids as acetic acid
    rAlkMgLcaco3 : REAL; // 碱度 [mg/L，以 CaCO3 计] / alkalinity as CaCO3
END_VAR
VAR_OUTPUT
    rRatio : REAL; // VFA/碱度比 [-] / VFA to alkalinity ratio
    bValid : BOOL; // 结果有效位 [-] / result valid flag
    iRisk : INT; // 风险等级 0=正常 1=关注 2=酸化预警 [-] / risk level
    iErrCode : INT; // 事件码 0=正常 1=碱度非法 2=比值超可观测上限 3=结果非有限 / event code
END_VAR
VAR CONSTANT
    rRiskWatch : REAL := 0.25; // 关注门槛 [-] / watch threshold
    rRiskAlarm : REAL := 0.4; // 酸化预警门槛 [-] / acidification alarm threshold
    rRatioCap : REAL := 100.0; // 比值输出饱和上限 [-] / ratio saturation cap
END_VAR
VAR
    rRatioRaw : REAL; // 未限幅比值 [-] / unchecked ratio
END_VAR

    // —— 段 0：全路径预清 —— //
    rRatioRaw := 0.0;
    rRatio := 0.0;
    iRisk := 0;
    bValid := FALSE;
    iErrCode := 0;
    FC_DL_VfaAlkalinityRatio := FALSE;
    // —— 段 1：分母闸（碱度必须为正） —— //
    IF rAlkMgLcaco3 <= 0.0 THEN
        iErrCode := 1; // 碱度非法，比值无定义 / invalid alkalinity, ratio undefined
        RETURN;
    END_IF;
    // —— 段 2：量纲链 (mg/L)/(mg/L) = 无量纲 —— //
    rRatioRaw := rVfaMgL / rAlkMgLcaco3; // 比值 [-] / ratio
    IF ABS(rRatioRaw) > 1.0E15 THEN
        iErrCode := 3; // 结果非有限，强制归零 / non-finite result, forced to zero
        RETURN;
    END_IF;
    // —— 段 3：负值防御与上限饱和 —— //
    IF rRatioRaw < 0.0 THEN
        rRatio := 0.0; // 负浓度防御 / negative concentration guard
    ELSIF rRatioRaw > rRatioCap THEN
        rRatio := rRatioCap; // 超上限饱和 / saturate at cap
        iErrCode := 2; // 信息级：比值超上限 / info level: ratio capped
    ELSE
        rRatio := rRatioRaw;
    END_IF;
    // —— 段 4：风险分级（用原始比值分级，避免饱和影响） —— //
    IF rRatioRaw > rRiskAlarm THEN
        iRisk := 2; // 酸化预警 / acidification alarm
    ELSIF rRatioRaw >= rRiskWatch THEN
        iRisk := 1; // 关注 / watch
    ELSE
        iRisk := 0; // 正常 / normal
    END_IF;
    bValid := TRUE;
    FC_DL_VfaAlkalinityRatio := TRUE;
END_FUNCTION

(* ---- FC_DL_WaterLangelierIndex.st ---- *)
(*
  ============================================================
  组件名 : FC_DL_WaterLangelierIndex
  分类   : DL_Process
  功能   : 水质朗格利尔饱和指数计算，由温度钙硬度碱度含盐量与 pH 判结垢或腐蚀倾向
  开源溯源 : internal-design（本轮无外部代码逐行引用）
             参考语义 : 无外部参考
  复杂度 : C2
  版本   : 1.0.0
  ============================================================
  口径说明 : A 为含盐量项 (log10(TDS)-1)/10，B 为温度项 -13.12*log10(T+273.15)+34.55，
             C 为钙硬度项 log10(CaHard)-0.4，D 为碱度项 log10(Alk)，pHs=(9.3+A+B)-(C+D)。
             本库 LOG 为十进制对数。指数大于 0.5 判结垢倾向，小于 -0.5 判腐蚀倾向。
*)

FUNCTION FC_DL_WaterLangelierIndex : REAL
VAR_INPUT
    rTempC      : REAL; // 水温 [摄氏度] water temperature [degree celsius]
    rCaHard_mgL : REAL; // 钙硬度（以碳酸钙计）[mg/L] calcium hardness as calcium carbonate [mg per litre]
    rAlk_mgL    : REAL; // 总碱度（以碳酸钙计）[mg/L] total alkalinity as calcium carbonate [mg per litre]
    rTds_mgL    : REAL; // 溶解性总固体 [mg/L] total dissolved solids [mg per litre]
    rPh         : REAL; // 实测 pH 值 [无量纲] measured pH value [dimensionless]
END_VAR
VAR_OUTPUT
    rLsi      : REAL; // 朗格利尔指数 [无量纲] Langelier saturation index [dimensionless]
    nTendency : INT; // 倾向 0平衡 1结垢 2腐蚀 [档] tendency 0 balanced, 1 scaling, 2 corrosive [band]
    rPhs      : REAL; // 饱和 pH 值 [无量纲] saturation pH value [dimensionless]
    bValid    : BOOL; // 结果有效标志 result validity flag
END_VAR
VAR CONSTANT
    DL_KELVIN    : REAL := 273.15; // 摄氏到开尔文偏移 celsius to kelvin offset
    DL_B_SLOPE   : REAL := 13.12; // 温度项斜率 the temperature term slope
    DL_B_OFFSET  : REAL := 34.55; // 温度项偏移 the temperature term offset
    DL_C_OFFSET  : REAL := 0.4; // 钙硬度项偏移 the calcium term offset
    DL_PHS_BASE  : REAL := 9.3; // 饱和 pH 基准常数 the saturation pH base constant
    DL_LSI_BAND  : REAL := 0.5; // 倾向判定带宽 [无量纲] tendency band [dimensionless]
    DL_TEN       : REAL := 10.0; // 含盐量项换算系数 the salinity term factor
    DL_EPS_R     : REAL := 1.0E-6; // 实数零判定阈值 real zero threshold
END_VAR
VAR
    _bFin : BOOL := FALSE; // 五输入有限性判定 finiteness verdict of the five inputs
    _rTempK : REAL := 0.0; // 绝对温度 [K] absolute temperature [K]
    _rA   : REAL := 0.0; // 含盐量项 [无量纲] salinity term [dimensionless]
    _rB   : REAL := 0.0; // 温度项 [无量纲] temperature term [dimensionless]
    _rC   : REAL := 0.0; // 钙硬度项 [无量纲] calcium term [dimensionless]
    _rD   : REAL := 0.0; // 碱度项 [无量纲] alkalinity term [dimensionless]
    _rPhs : REAL := 0.0; // 饱和 pH 中间量 [无量纲] intermediate saturation pH [dimensionless]
    _rLsi : REAL := 0.0; // 指数中间量 [无量纲] intermediate index [dimensionless]
END_VAR

// 段 1｜出口预置 preset the exit
FC_DL_WaterLangelierIndex := 0.0; // 缺省返回零 default zero return
rLsi := 0.0; // 指数预置零 index preset to zero
nTendency := 0; // 倾向预置平衡 tendency preset balanced
rPhs := 0.0; // 饱和 pH 预置零 saturation pH preset to zero
bValid := FALSE; // 计算完成前不认结果 unusable before the calculation
// 段 2｜非有限闸 finiteness gate
_bFin := (rTempC = rTempC) AND (rCaHard_mgL = rCaHard_mgL) AND (rAlk_mgL = rAlk_mgL) AND (rTds_mgL = rTds_mgL) AND (rPh = rPh); // 五输入自反判定 self comparison of the five inputs
IF NOT _bFin THEN
    RETURN; // 非有限即无效 non finite means invalid
END_IF
// 段 3｜取对数项的正值闸 positive value gate for the logarithm terms
IF (rCaHard_mgL <= DL_EPS_R) OR (rAlk_mgL <= DL_EPS_R) OR (rTds_mgL <= DL_EPS_R) THEN
    RETURN; // 浓度非正无法取对数 a non positive concentration cannot carry a logarithm
END_IF
_rTempK := rTempC + DL_KELVIN; // 摄氏折算绝对温度 celsius to absolute temperature
IF _rTempK <= DL_EPS_R THEN
    RETURN; // 绝对温度非正无法取对数 a non positive absolute temperature cannot carry a logarithm
END_IF
// 段 4｜四项折算与饱和 pH the four terms and the saturation pH
_rA := (LOG(rTds_mgL) - 1.0) / DL_TEN; // 含盐量项 salinity term
_rB := 0.0 - DL_B_SLOPE * LOG(_rTempK) + DL_B_OFFSET; // 温度项 temperature term
_rC := LOG(rCaHard_mgL) - DL_C_OFFSET; // 钙硬度项 calcium hardness term
_rD := LOG(rAlk_mgL); // 碱度项 alkalinity term
_rPhs := (DL_PHS_BASE + _rA + _rB) - (_rC + _rD); // 饱和 pH saturation pH
rPhs := _rPhs; // 饱和 pH 落定 land the saturation pH
// 段 5｜指数与倾向判定 index and the tendency verdict
_rLsi := rPh - _rPhs; // 实测 pH 减饱和 pH measured minus the saturation value
rLsi := _rLsi; // 指数落定 land the index
IF _rLsi > DL_LSI_BAND THEN
    nTendency := 1; // 结垢倾向 scaling tendency
ELSIF _rLsi < (0.0 - DL_LSI_BAND) THEN
    nTendency := 2; // 腐蚀倾向 corrosive tendency
ELSE
    nTendency := 0; // 基本平衡 nearly balanced
END_IF
bValid := TRUE; // 结果可用 result usable
FC_DL_WaterLangelierIndex := _rLsi; // 函数返回指数 return the index
END_FUNCTION

(* ---- FC_DL_WaterRecoveryRatio.st ---- *)
(*
  ============================================================
  组件名 : FC_DL_WaterRecoveryRatio
  分类   : DL_Process
  功能   : 水处理系统回收率计算，含进料产水浓水三流股的物料平衡校核
  开源溯源 : internal-design（本轮无外部代码逐行引用）
             参考语义 : 无外部参考
  复杂度 : C1
  版本   : 1.0.0
  ============================================================
*)

FUNCTION FC_DL_WaterRecoveryRatio : REAL
VAR_INPUT
    rPermeate_m3h        : REAL; // 产水流量 [m3/h] permeate flow [m3 per hour]
    rFeed_m3h            : REAL; // 进料流量 [m3/h] feed flow [m3 per hour]
    rConc_m3h            : REAL; // 浓水流量 [m3/h] concentrate flow [m3 per hour]
    bCheckMassBalance    : BOOL; // 真为启用物料平衡校核 enable the mass balance check when true
END_VAR
VAR_OUTPUT
    rRecoveryPct  : REAL; // 回收率 [%] recovery percentage [%]
    rMassBalErrPct: REAL; // 物料平衡偏差 [%] mass balance error [%]
    bValid        : BOOL; // 结果有效标志 result validity flag
END_VAR
VAR CONSTANT
    DL_HUNDRED   : REAL := 100.0; // 百分制换算系数 percentage scale factor
    DL_BAL_LIMIT : REAL := 5.0; // 物料平衡允许偏差 [%] admissible balance error [%]
    DL_EPS_R     : REAL := 1.0E-6; // 实数零判定阈值 real zero threshold
END_VAR
VAR
    _bFin : BOOL := FALSE; // 三实数输入有限性判定 finiteness verdict of the three real inputs
    _rRec : REAL := 0.0; // 回收率中间量 [%] intermediate recovery [%]
    _rBal : REAL := 0.0; // 平衡偏差中间量 [%] intermediate balance error [%]
END_VAR

// 段 1｜出口预置 preset the exit
FC_DL_WaterRecoveryRatio := 0.0; // 缺省返回零 default zero return
rRecoveryPct := 0.0; // 回收率预置零 recovery preset to zero
rMassBalErrPct := 0.0; // 平衡偏差预置零 balance error preset to zero
bValid := FALSE; // 计算完成前不认结果 unusable before the calculation
// 段 2｜非有限闸 finiteness gate
_bFin := (rPermeate_m3h = rPermeate_m3h) AND (rFeed_m3h = rFeed_m3h) AND (rConc_m3h = rConc_m3h); // 三输入自反判定 self comparison of the three inputs
IF NOT _bFin THEN
    RETURN; // 非有限即无效 non finite means invalid
END_IF
// 段 3｜进料分母闸与负流量闸 feed divisor gate and negative flow gate
IF rFeed_m3h <= DL_EPS_R THEN
    RETURN; // 进料非正无法折算回收率 a non positive feed cannot carry a recovery
END_IF
IF (rPermeate_m3h < 0.0) OR (rConc_m3h < 0.0) THEN
    RETURN; // 负流量属采集异常 a negative flow is a measurement fault
END_IF
// 段 4｜回收率与物料平衡 recovery and the mass balance
_rRec := rPermeate_m3h / rFeed_m3h * DL_HUNDRED; // 产水占进料百分比 permeate over feed as a percentage
_rBal := (rFeed_m3h - rPermeate_m3h - rConc_m3h) / rFeed_m3h * DL_HUNDRED; // 三流股闭合偏差 closure error of the three streams
rRecoveryPct := _rRec; // 回收率落定 land the recovery
rMassBalErrPct := _rBal; // 平衡偏差落定 land the balance error
// 段 5｜按需物料平衡校核 conditional mass balance check
IF bCheckMassBalance AND (ABS(_rBal) > DL_BAL_LIMIT) THEN
    RETURN; // 平衡超差判无效 an excessive balance error is void
END_IF
bValid := TRUE; // 结果可用 result usable
FC_DL_WaterRecoveryRatio := _rRec; // 函数返回回收率 return the recovery
END_FUNCTION

(* ---- FC_DL_WeighBatchYieldCalc.st ---- *)
(*
  ============================================================
  组件名 : FC_DL_WeighBatchYieldCalc
  分类   : DL_Process
  功能   : 批次实际投料与理论投料的收得率百分比计算与公差判定
  开源溯源 : internal-design（本轮无外部代码逐行引用）
             参考语义 : 无外部参考
  复杂度 : C1
  版本   : 1.0.0
  ============================================================
*)

FUNCTION FC_DL_WeighBatchYieldCalc : REAL
VAR_INPUT
    rActualFeed  : REAL; // 实际投料量 [kg] actual feed quantity [kg]
    rTheoryFeed  : REAL; // 理论投料量 [kg] theoretical feed quantity [kg]
    rTolPct      : REAL; // 收得率公差 [%] yield tolerance [%]
END_VAR
VAR_OUTPUT
    rYieldPct : REAL; // 收得率 [%] yield percentage [%]
    bInTol    : BOOL; // 收得率在公差内标志 yield inside tolerance flag
    bValid    : BOOL; // 结果有效标志 result validity flag
END_VAR
VAR CONSTANT
    DL_EPS_R : REAL := 1.0E-6; // 实数零判定阈值 real zero threshold
    DL_HUNDRED : REAL := 100.0; // 百分制换算系数 percentage scale factor
END_VAR
VAR
    _bFin : BOOL := FALSE; // 两实数输入有限性判定 finiteness verdict of both real inputs
    _rTol : REAL := 0.0; // 钳位后的公差 [%] clamped tolerance [%]
END_VAR

// 段 1｜出口预置 preset the exit
FC_DL_WeighBatchYieldCalc := 0.0; // 缺省返回零 default zero return
rYieldPct := 0.0; // 收得率预置零 yield preset to zero
bInTol := FALSE; // 公差内标志预置假 tolerance flag preset false
bValid := FALSE; // 计算完成前不认结果 unusable before the calculation
// 段 2｜非有限闸 finiteness gate
_bFin := (rActualFeed = rActualFeed) AND (rTheoryFeed = rTheoryFeed) AND (rTolPct = rTolPct); // 三输入自反判定 self comparison of the three inputs
IF NOT _bFin THEN
    RETURN; // 非有限即无效 non finite means invalid
END_IF
// 段 3｜理论投料量分母闸 theoretical feed divisor gate
IF rTheoryFeed <= DL_EPS_R THEN
    RETURN; // 理论量非正无法折算收得率 a non positive theory cannot carry a yield
END_IF
// 段 4｜收得率与公差判定 yield computation and the tolerance verdict
rYieldPct := rActualFeed / rTheoryFeed * DL_HUNDRED; // 收得率百分比 yield percentage
_rTol := rTolPct; // 取入参公差 take the tolerance input
IF _rTol < 0.0 THEN
    _rTol := ABS(_rTol); // 负公差取幅值 a negative tolerance becomes its magnitude
END_IF
bInTol := ABS(rYieldPct - DL_HUNDRED) <= _rTol; // 对百分之百的双向公差带 symmetric tolerance band around one hundred percent
bValid := TRUE; // 结果可用 result usable
FC_DL_WeighBatchYieldCalc := rYieldPct; // 函数返回收得率 return the yield
END_FUNCTION

(* ---- FC_DL_WeighCreepCompensate.st ---- *)
(*
  ============================================================
  组件名 : FC_DL_WeighCreepCompensate
  分类   : DL_Process
  功能   : 称重传感器蠕变补偿，按加载时长、蠕变速率与温度因子修正原始读数
  开源溯源 : internal-design（本轮无外部代码逐行引用）
             参考语义 : 无外部参考
  复杂度 : C1
  版本   : 1.0.0
  ============================================================
*)

FUNCTION FC_DL_WeighCreepCompensate : REAL
VAR_INPUT
    rRaw              : REAL; // 传感器原始读数 [kg] raw load cell reading [kg]
    rLoadTimeS        : REAL; // 持续加载时长 [s] continuous loaded duration [s]
    rCreepRatePctPerH : REAL; // 每小时蠕变百分比 [%/h] creep percentage per hour [%/h]
    rTempFactor       : REAL; // 温度修正因子 1.0 为常温 [无量纲] temperature factor, one at ambient [dimensionless]
END_VAR
VAR_OUTPUT
    rCorrected : REAL; // 蠕变补偿后的读数 [kg] creep corrected reading [kg]
    bValid     : BOOL; // 结果有效标志 result validity flag
END_VAR
VAR CONSTANT
    DL_SEC_PER_HOUR : REAL := 3600.0; // 每小时秒数 seconds per hour
    DL_HUNDRED      : REAL := 100.0; // 百分制换算系数 percentage scale factor
END_VAR
VAR
    _bFin  : BOOL := FALSE; // 四输入有限性判定 finiteness verdict of the four inputs
    _rRel  : REAL := 0.0; // 累计相对蠕变量 [无量纲] accumulated relative creep [dimensionless]
    _rCorr : REAL := 0.0; // 修正后的读数中间量 [kg] intermediate corrected reading [kg]
END_VAR

// 段 1｜出口预置 preset the exit
FC_DL_WeighCreepCompensate := 0.0; // 缺省返回零 default zero return
rCorrected := 0.0; // 修正值预置零 corrected value preset to zero
bValid := FALSE; // 计算完成前不认结果 unusable before the calculation
// 段 2｜非有限闸 finiteness gate
_bFin := (rRaw = rRaw) AND (rLoadTimeS = rLoadTimeS) AND (rCreepRatePctPerH = rCreepRatePctPerH) AND (rTempFactor = rTempFactor); // 四输入自反判定 self comparison of the four inputs
IF NOT _bFin THEN
    RETURN; // 非有限即无效 non finite means invalid
END_IF
// 段 3｜时长与速率方向闸 duration and rate direction gate
IF (rLoadTimeS < 0.0) OR (rCreepRatePctPerH < 0.0) THEN
    RETURN; // 负时长或负速率属配置非法 a negative duration or rate is an illegal configuration
END_IF
// 段 4｜蠕变量折算与主体补偿 creep quantity and the main compensation
_rRel := rCreepRatePctPerH / DL_HUNDRED * (rLoadTimeS / DL_SEC_PER_HOUR) * rTempFactor; // 相对蠕变量 relative creep quantity
_rCorr := rRaw * (1.0 + _rRel); // 原始读数按蠕变量放大 amplify the raw reading by the creep quantity
IF (_rCorr <> _rCorr) OR (ABS(_rCorr) > 1.0E30) THEN
    RETURN; // 结果非有限拒收 refuse a non finite result
END_IF
rCorrected := _rCorr; // 修正值落定 land the corrected value
bValid := TRUE; // 结果可用 result usable
FC_DL_WeighCreepCompensate := _rCorr; // 函数返回修正值 return the corrected value
END_FUNCTION

(* ---- FC_DL_WeighDoseTolBand.st ---- *)
(*
  ============================================================
  组件名 : FC_DL_WeighDoseTolBand
  分类   : DL_Process
  功能   : 配料实绩对目标值的公差带判定，返回欠量、合格、超量或无效分档
  开源溯源 : internal-design（本轮无外部代码逐行引用）
             参考语义 : 无外部参考
  复杂度 : C1
  版本   : 1.0.0
  ============================================================
*)

FUNCTION FC_DL_WeighDoseTolBand : INT
VAR_INPUT
    rTarget      : REAL; // 配料目标值 [kg] dosing target [kg]
    rActual      : REAL; // 配料实绩值 [kg] actual dosed weight [kg]
    rTolMinus    : REAL; // 下公差（欠量侧）[kg] minus tolerance on the under side [kg]
    rTolPlus     : REAL; // 上公差（超量侧）[kg] plus tolerance on the over side [kg]
    rMinEffective: REAL; // 有效称量下限 [kg] minimum effective reading [kg]
END_VAR
VAR_OUTPUT
    nBand  : INT; // 分档结果 -2无效 -1欠 0合格 1超 [档] band code -2 void, -1 under, 0 ok, 1 over [band]
    bValid : BOOL; // 结果有效标志 result validity flag
END_VAR
VAR
    _bFin  : BOOL := FALSE; // 三实数输入有限性判定 finiteness verdict of the three real inputs
    _rTolM : REAL := 0.0; // 钳位后的下公差 [kg] clamped minus tolerance [kg]
    _rTolP : REAL := 0.0; // 钳位后的上公差 [kg] clamped plus tolerance [kg]
    _rLow  : REAL := 0.0; // 合格带下沿 [kg] lower edge of the band [kg]
    _rHigh : REAL := 0.0; // 合格带上沿 [kg] upper edge of the band [kg]
END_VAR

// 段 1｜出口预置 preset the exit
FC_DL_WeighDoseTolBand := -2; // 缺省按无效分档 default void band
nBand := -2; // 分档码预置无效 band code preset void
bValid := FALSE; // 计算完成前不认结果 unusable before the calculation
// 段 2｜非有限闸 finiteness gate
_bFin := (rTarget = rTarget) AND (rActual = rActual) AND (rTolMinus = rTolMinus) AND (rTolPlus = rTolPlus) AND (rMinEffective = rMinEffective); // 五输入自反判定 self comparison of the five inputs
IF NOT _bFin THEN
    RETURN; // 非有限即无效 non finite means invalid
END_IF
// 段 3｜有效称量下限闸 minimum effective reading gate
IF rActual < rMinEffective THEN
    RETURN; // 读数低于有效下限按无效处理 a reading below the floor is void
END_IF
// 段 4｜公差整形与带沿计算 tolerance reshape and band edges
_rTolM := rTolMinus; // 取下公差 take the minus tolerance
IF _rTolM < 0.0 THEN
    _rTolM := ABS(_rTolM); // 负下公差取幅值 a negative minus tolerance becomes its magnitude
END_IF
_rTolP := rTolPlus; // 取上公差 take the plus tolerance
IF _rTolP < 0.0 THEN
    _rTolP := ABS(_rTolP); // 负上公差取幅值 a negative plus tolerance becomes its magnitude
END_IF
_rLow := rTarget - _rTolM; // 合格带下沿 lower edge of the acceptance band
_rHigh := rTarget + _rTolP; // 合格带上沿 upper edge of the acceptance band
// 段 5｜双向分档判定 directional band verdict
IF rActual < _rLow THEN
    nBand := -1; // 欠量 under weight
ELSIF rActual > _rHigh THEN
    nBand := 1; // 超量 over weight
ELSE
    nBand := 0; // 带内合格 in band
END_IF
bValid := TRUE; // 结果可用 result usable
FC_DL_WeighDoseTolBand := nBand; // 函数返回分档码 return the band code
END_FUNCTION

(* ---- FC_DL_WeighMultiHeadSum.st ---- *)
(*
  ============================================================
  组件名 : FC_DL_WeighMultiHeadSum
  分类   : DL_Process
  功能   : 多头组合称重穷举，选出不低于目标欠量下限且偏差最小的头组合位图
  开源溯源 : internal-design（本轮无外部代码逐行引用）
             参考语义 : 无外部参考
  复杂度 : C2
  版本   : 1.0.0
  ============================================================
*)

FUNCTION FC_DL_WeighMultiHeadSum : REAL
VAR_INPUT
    aWeight   : ARRAY[0..7] OF REAL; // 八只称重头实测值 [kg] measured weights of eight heads [kg]
    nHeads    : INT; // 参与组合的头数 1~8 [个] engaged head count from one to eight [count]
    rTarget   : REAL; // 目标组合重量 [kg] target combination weight [kg]
    rAllowTol : REAL; // 允许欠量容差 [kg] allowed under weight tolerance [kg]
END_VAR
VAR_OUTPUT
    rBestSum   : REAL; // 最优组合和 [kg] best combination sum [kg]
    nBestMask  : INT; // 最优组合位图 [位图] best combination bit mask [bit map]
    nBestCount : INT; // 最优组合头数 [个] head count of the best combination [count]
    bValid     : BOOL; // 结果有效标志 result validity flag
END_VAR
VAR
    nMask  : INT := 0; // 组合位图游标 [位图] combination mask cursor [bit map]
    nBit   : INT := 0; // 位游标 0~7 [位] bit cursor from zero to seven [bit]
    nRem   : INT := 0; // 位图右移余量 [位图] mask remainder while shifting [bit map]
    nCnt   : INT := 0; // 当前组合头数 [个] head count of the current mask [count]
    rSum   : REAL := 0.0; // 当前组合和 [kg] sum of the current mask [kg]
    rBest  : REAL := 0.0; // 当前最优组合和 [kg] best sum found so far [kg]
    rErr   : REAL := 0.0; // 当前组合偏差绝对值 [kg] absolute deviation of the current mask [kg]
    rMin   : REAL := 0.0; // 当前最小偏差绝对值 [kg] smallest absolute deviation so far [kg]
    rFloor : REAL := 0.0; // 允许的组合和下限 [kg] lower admissible sum [kg]
    bHit   : BOOL := FALSE; // 找到候选组合标志 candidate found flag
    _bFin  : BOOL := FALSE; // 实数输入有限性判定 finiteness verdict of the real inputs
END_VAR

// 段 1｜出口预置 preset the exit
FC_DL_WeighMultiHeadSum := 0.0; // 缺省返回零 default zero return
rBestSum := 0.0; // 最优和预置零 best sum preset to zero
nBestMask := 0; // 位图预置零 bit mask preset to zero
nBestCount := 0; // 头数预置零 head count preset to zero
bValid := FALSE; // 计算完成前不认结果 unusable before the calculation
// 段 2｜头数闸与有限闸 head count gate and finiteness gate
_bFin := (rTarget = rTarget) AND (rAllowTol = rAllowTol); // 两实数输入自反判定 self comparison of both real inputs
IF (NOT _bFin) OR (nHeads < 1) OR (nHeads > 8) THEN
    RETURN; // 头数越界或非有限即无效 an out of range head count or a non finite input is void
END_IF
rFloor := rTarget - ABS(rAllowTol); // 允许下限取容差幅值 the floor uses the tolerance magnitude
// 段 3｜穷举 255 个非零组合 exhaustive walk of two hundred fifty five non empty masks
FOR nMask := 1 TO 255 DO
    nCnt := 0; // 组合头数清零 clear the head count
    rSum := 0.0; // 组合和清零 clear the sum
    nRem := nMask; // 余量取位图 the remainder starts from the mask
    FOR nBit := 0 TO 7 DO
        IF ((nRem MOD 2) = 1) AND (nBit < nHeads) THEN
            nCnt := nCnt + 1; // 头数累加 accumulate the head count
            rSum := rSum + aWeight[nBit]; // 重量累加 accumulate the weight
        END_IF
        nRem := nRem / 2; // 整数除二右移一位 integer division by two shifts one bit
    END_FOR
    // 段 4｜候选判据与最优保持 candidate verdict and the best hold
    IF (nCnt > 0) AND (rSum >= rFloor) THEN
        rErr := ABS(rSum - rTarget); // 组合偏差绝对值 absolute deviation of the mask
        IF (NOT bHit) OR (rErr < rMin) THEN
            rMin := rErr; // 更新最小偏差 refresh the smallest deviation
            rBest := rSum; // 更新最优组合和 refresh the best sum
            nBestMask := nMask; // 更新最优位图 refresh the best mask
            nBestCount := nCnt; // 更新最优头数 refresh the best head count
            bHit := TRUE; // 置候选命中标志 raise the candidate flag
        END_IF
    END_IF
END_FOR
// 段 5｜出口与命中判定 the exit and the hit verdict
IF bHit THEN
    rBestSum := rBest; // 最优和落定 land the best sum
    bValid := TRUE; // 结果可用 result usable
    FC_DL_WeighMultiHeadSum := rBest; // 函数返回最优和 return the best sum
END_IF
END_FUNCTION

(* ---- FC_DL_WeighNetFromGross.st ---- *)
(*
  ============================================================
  组件名 : FC_DL_WeighNetFromGross
  分类   : DL_Process
  功能   : 毛重去皮与零点偏置扣除求净重，负净重超出容差判无效并清零
  开源溯源 : internal-design（本轮无外部代码逐行引用）
             参考语义 : 无外部参考
  复杂度 : C1
  版本   : 1.0.0
  ============================================================
*)

FUNCTION FC_DL_WeighNetFromGross : REAL
VAR_INPUT
    rGross      : REAL; // 毛重 [kg] gross weight [kg]
    rTare       : REAL; // 皮重 [kg] tare weight [kg]
    rZeroOffset : REAL; // 零点偏置 [kg] zero offset [kg]
    rNegTol     : REAL; // 负净重容差 [kg] negative net tolerance [kg]
END_VAR
VAR_OUTPUT
    rNet   : REAL; // 净重结果 [kg] net weight result [kg]
    bValid : BOOL; // 结果有效标志 result validity flag
END_VAR
VAR
    _bFin : BOOL := FALSE; // 四输入有限性判定 finiteness verdict of the four inputs
    _rTol : REAL := 0.0; // 钳位后的负容差 [kg] clamped negative tolerance [kg]
    _rNet : REAL := 0.0; // 净重中间量 [kg] intermediate net weight [kg]
END_VAR

// 段 1｜出口预置 preset the exit
FC_DL_WeighNetFromGross := 0.0; // 缺省返回零 default zero return
rNet := 0.0; // 净重预置零 net weight preset to zero
bValid := FALSE; // 计算完成前不认结果 unusable before the calculation
// 段 2｜非有限闸 finiteness gate
_bFin := (rGross = rGross) AND (rTare = rTare) AND (rZeroOffset = rZeroOffset) AND (rNegTol = rNegTol); // 四输入自反判定 self comparison of the four inputs
IF NOT _bFin THEN
    RETURN; // 非有限即无效，出口保持零点 non finite means invalid and the zero output stays
END_IF
// 段 3｜负容差整形 reshape the negative tolerance
_rTol := rNegTol; // 取入参容差 take the tolerance input
IF _rTol < 0.0 THEN
    _rTol := 0.0; // 负容差按零处理 a negative tolerance becomes zero
END_IF
// 段 4｜主体扣减与负净重拦截 main subtraction and the negative net gate
_rNet := rGross - rTare - rZeroOffset; // 毛重去皮去零点 gross minus tare minus zero offset
IF _rNet < -_rTol THEN
    rNet := 0.0; // 超负容差净重清零 clear the net weight beyond tolerance
    RETURN; // 判无效并早退 invalid and early return
END_IF
rNet := _rNet; // 净重落定 land the net weight
bValid := TRUE; // 结果可用 result usable
FC_DL_WeighNetFromGross := _rNet; // 函数返回净重 return the net weight
END_FUNCTION
